FUNCTION "FRK_PersistCommitAnchor" : Void
{ S7_Optimized_Access := 'TRUE' }
VERSION : 0.1
VAR_INPUT
    Slot : Int;
END_VAR
BEGIN
    IF #Slot < 1 OR #Slot > 18 THEN RETURN; END_IF;
    IF "FRK_PersistAnchors".SelectedB[#Slot] THEN "FRK_PersistAnchors".RowsA[#Slot] := "FRK_PersistRuntime".Anchor[#Slot];
    ELSE "FRK_PersistAnchors".RowsB[#Slot] := "FRK_PersistRuntime".Anchor[#Slot]; END_IF;
    "FRK_PersistAnchors".SelectedB[#Slot] := NOT "FRK_PersistAnchors".SelectedB[#Slot];
    "FRK_PersistAnchors".Commissioned[#Slot] := TRUE;
END_FUNCTION
// Binding-owned byte medium. Consumers own content validation and authority.
FUNCTION "FRK_PersistNumber" : DWord
{ S7_Optimized_Access := 'TRUE' }
VERSION : 0.1
VAR_INPUT
    Offset : Int;
END_VAR
VAR_IN_OUT
    Bytes : Array[*] of Byte;
END_VAR
VAR_TEMP
    Index : Int;
END_VAR
BEGIN
    #FRK_PersistNumber := DWORD#0;
    IF #Offset < 0 OR #Offset > UPPER_BOUND(ARR := #Bytes, DIM := 1) - 3 THEN RETURN; END_IF;
    FOR #Index := 0 TO 3 DO
        #FRK_PersistNumber := #FRK_PersistNumber OR SHL(IN := BYTE_TO_DWORD(#Bytes[#Offset + #Index]), N := INT_TO_UINT(#Index * 8));
    END_FOR;
END_FUNCTION

FUNCTION "FRK_PersistPutNumber" : Void
{ S7_Optimized_Access := 'TRUE' }
VERSION : 0.1
VAR_INPUT
    Offset : Int;
    Value : DWord;
END_VAR
VAR_IN_OUT
    Bytes : Array[*] of Byte;
END_VAR
VAR_TEMP
    Index : Int;
END_VAR
BEGIN
    IF #Offset < 0 OR #Offset > UPPER_BOUND(ARR := #Bytes, DIM := 1) - 3 THEN RETURN; END_IF;
    FOR #Index := 0 TO 3 DO #Bytes[#Offset + #Index] := DWORD_TO_BYTE(SHR(IN := #Value, N := INT_TO_UINT(#Index * 8))); END_FOR;
END_FUNCTION

FUNCTION "FRK_PersistKeyCrc" : DWord
{ S7_Optimized_Access := 'TRUE' }
VERSION : 0.1
VAR_INPUT
    Key : String;
END_VAR
VAR_TEMP
    Index : Int;
    Work : DWord;
END_VAR
BEGIN
    #Work := "FRK_CrcNumber"(Previous := DWORD#16#FFFFFFFF, Value := INT_TO_UDINT(LEN(#Key)));
    FOR #Index := 1 TO LEN(#Key) DO #Work := "FRK_CrcByte"(Previous := #Work, Value := CHAR_TO_BYTE(#Key[#Index])); END_FOR;
    #FRK_PersistKeyCrc := NOT #Work;
END_FUNCTION

FUNCTION "FRK_PersistAnchorCrc" : DWord
{ S7_Optimized_Access := 'TRUE' }
VERSION : 0.1
VAR_IN_OUT
    Image : "FRK_PersistAnchor";
END_VAR
VAR_TEMP
    Work : DWord;
END_VAR
BEGIN
    #Work := "FRK_CrcNumber"(Previous := DWORD#16#FFFFFFFF, Value := UINT_TO_UDINT(#Image.SchemaVersion));
    #Work := "FRK_CrcNumber"(Previous := #Work, Value := DWORD_TO_UDINT(#Image.KeyCrc));
    #Work := "FRK_CrcNumber"(Previous := #Work, Value := #Image.Generation);
    #Work := "FRK_CrcNumber"(Previous := #Work, Value := DWORD_TO_UDINT(#Image.DocumentCrc));
    #FRK_PersistAnchorCrc := NOT #Work;
END_FUNCTION

FUNCTION "FRK_PersistAnchorValid" : Bool
{ S7_Optimized_Access := 'TRUE' }
VERSION : 0.1
VAR_INPUT
    Slot : Int;
END_VAR
BEGIN
    #FRK_PersistAnchorValid := FALSE;
    IF #Slot < 1 OR #Slot > 18 THEN RETURN; END_IF;
    #FRK_PersistAnchorValid := "FRK_PersistAnchors".Commissioned[#Slot]
        AND "FRK_PersistRuntime".Anchor[#Slot].SchemaVersion = 1
        AND "FRK_PersistRuntime".Anchor[#Slot].KeyCrc = "FRK_PersistRuntime".KeyCrc[#Slot]
        AND "FRK_PersistRuntime".Anchor[#Slot].Checksum = "FRK_PersistAnchorCrc"(Image := "FRK_PersistRuntime".Anchor[#Slot]);
END_FUNCTION

FUNCTION "FRK_PersistRepair" : Void
{ S7_Optimized_Access := 'TRUE' }
VERSION : 0.1
VAR_INPUT
    Slot : Int;
END_VAR
BEGIN
    // Trusted consumer seam; never a remote command or authorization authority.
    IF #Slot < 1 OR #Slot > 18 THEN RETURN; END_IF;
    IF NOT "FRK_PersistAnchorValid"(Slot := #Slot) THEN
        "FRK_PersistRuntime".Anchor[#Slot].SchemaVersion := 1;
        "FRK_PersistRuntime".Anchor[#Slot].KeyCrc := "FRK_PersistRuntime".KeyCrc[#Slot];
        "FRK_PersistRuntime".Anchor[#Slot].Generation := 0;
        "FRK_PersistRuntime".Anchor[#Slot].DocumentCrc := DWORD#0;
        "FRK_PersistRuntime".Anchor[#Slot].Checksum := "FRK_PersistAnchorCrc"(Image := "FRK_PersistRuntime".Anchor[#Slot]);
        "FRK_PersistAnchors".Commissioned[#Slot] := TRUE;
    END_IF;
    "FRK_PersistCommitAnchor"(Slot := #Slot);
END_FUNCTION

FUNCTION "FRK_PersistStart" : UDInt
{ S7_Optimized_Access := 'TRUE' }
VERSION : 0.1
VAR_INPUT
    Slot : Int;
    WriteDocument : Bool;
    Length : DInt;
END_VAR
VAR_TEMP
    Index : Int;
END_VAR
BEGIN
    #FRK_PersistStart := 0;
    IF #Slot < 1 OR #Slot > 18 THEN RETURN; END_IF;
    IF #Length < 0 OR #Length > "FRK_PersistRuntime".Capacity[#Slot] OR "FRK_PersistRuntime".Leased[#Slot] THEN RETURN; END_IF;
    IF "FRK_PersistRuntime".LastTicket = UDINT#4294967295 THEN RETURN; END_IF;
    FOR #Index := 1 TO 4 DO
        IF "FRK_PersistRuntime".Queue[#Index].State = 0 THEN
            "FRK_PersistRuntime".LastTicket := "FRK_PersistRuntime".LastTicket + 1;
            "FRK_PersistRuntime".Queue[#Index].Ticket := "FRK_PersistRuntime".LastTicket;
            "FRK_PersistRuntime".Queue[#Index].Slot := #Slot;
            "FRK_PersistRuntime".Queue[#Index].WriteDocument := #WriteDocument;
            "FRK_PersistRuntime".Queue[#Index].Length := #Length;
            "FRK_PersistRuntime".Queue[#Index].State := 1;
            "FRK_PersistRuntime".Leased[#Slot] := TRUE;
            #FRK_PersistStart := "FRK_PersistRuntime".LastTicket;
            RETURN;
        END_IF;
    END_FOR;
END_FUNCTION

FUNCTION "FRK_PersistFinish" : Void
{ S7_Optimized_Access := 'TRUE' }
VERSION : 0.1
BEGIN
    IF "FRK_PersistRuntime".Active < 1 OR "FRK_PersistRuntime".Active > 4 THEN RETURN; END_IF;
    "FRK_PersistRuntime".Queue["FRK_PersistRuntime".Active].Result := "FRK_PersistRuntime".Result;
    "FRK_PersistRuntime".Queue["FRK_PersistRuntime".Active].State := 3;
    "FRK_PersistRuntime".Active := 0;
    "FRK_PersistRuntime".Stage := 0;
END_FUNCTION

FUNCTION "FRK_PersistValidate" : Bool
{ S7_Optimized_Access := 'TRUE' }
VERSION : 0.1
VAR_INPUT
    ExpectedKey : DWord;
END_VAR
VAR_IN_OUT
    Bytes : Array[*] of Byte;
    Check : "FRK_PersistCheck";
END_VAR
VAR_TEMP
    Budget : Int;
    Offset : Int;
    Upper : Int;
END_VAR
BEGIN
    #FRK_PersistValidate := FALSE;
    #Upper := DINT_TO_INT(UPPER_BOUND(ARR := #Bytes, DIM := 1));
    IF #Check.Cursor = -1 THEN
        #Check.Valid := FALSE; #Check.Empty := TRUE; #Check.Generation := 0; #Check.Length := 0;
        #Check.Cursor := 0; #Check.Crc := DWORD#16#FFFFFFFF;
        #Check.ZeroMode := "FRK_PersistNumber"(Offset := 0, Bytes := #Bytes) = DWORD#0;
        IF NOT #Check.ZeroMode THEN
            #Check.Empty := FALSE;
            IF "FRK_PersistNumber"(Offset := 0, Bytes := #Bytes) <> DWORD#826559046
                OR "FRK_PersistNumber"(Offset := 4, Bytes := #Bytes) <> DWORD#1
                OR "FRK_PersistNumber"(Offset := 16, Bytes := #Bytes) <> #ExpectedKey THEN #FRK_PersistValidate := TRUE; RETURN; END_IF;
            #Check.Generation := DWORD_TO_UDINT("FRK_PersistNumber"(Offset := 8, Bytes := #Bytes));
            #Check.Length := DWORD_TO_UDINT("FRK_PersistNumber"(Offset := 12, Bytes := #Bytes));
            IF #Check.Generation = 0 OR #Check.Length > INT_TO_UDINT(#Upper + 1 - 24) THEN #FRK_PersistValidate := TRUE; RETURN; END_IF;
        END_IF;
    END_IF;
    #Budget := 0;
    IF #Check.ZeroMode THEN
        WHILE #Check.Cursor <= #Upper AND #Budget < 512 DO
            IF #Bytes[#Check.Cursor] <> BYTE#0 THEN #Check.Empty := FALSE; #FRK_PersistValidate := TRUE; RETURN; END_IF;
            #Check.Cursor := #Check.Cursor + 1; #Budget := #Budget + 1;
        END_WHILE;
        #FRK_PersistValidate := #Check.Cursor > #Upper;
    ELSE
        WHILE #Check.Cursor < 20 + UDINT_TO_DINT(#Check.Length) AND #Budget < 512 DO
            IF #Check.Cursor < 20 THEN #Offset := DINT_TO_INT(#Check.Cursor); ELSE #Offset := DINT_TO_INT(#Check.Cursor + 24 - 20); END_IF;
            #Check.Crc := "FRK_CrcByte"(Previous := #Check.Crc, Value := #Bytes[#Offset]);
            #Check.Cursor := #Check.Cursor + 1; #Budget := #Budget + 1;
        END_WHILE;
        IF #Check.Cursor >= 20 + UDINT_TO_DINT(#Check.Length) THEN
            #Check.Crc := NOT #Check.Crc;
            #Check.Valid := #Check.Crc = "FRK_PersistNumber"(Offset := 20, Bytes := #Bytes);
            #FRK_PersistValidate := TRUE;
        END_IF;
    END_IF;
END_FUNCTION

FUNCTION "FRK_PersistInspect" : Void
{ S7_Optimized_Access := 'TRUE' }
VERSION : 0.1
VAR_IN_OUT
    BytesA : Array[*] of Byte;
    BytesB : Array[*] of Byte;
    Payload : Array[*] of Byte;
END_VAR
VAR_TEMP
    Index : Int;
    Slot : Int;
    Chosen : Int;
    Generation : UDInt;
    Length : UDInt;
    DocumentCrc : DWord;
    Lost : Bool;
END_VAR
BEGIN
    #Slot := "FRK_PersistRuntime".Slot;
    #Chosen := 0; #Generation := 0; #Length := 0; #DocumentCrc := DWORD#0;
    IF "FRK_PersistRuntime".CheckA.Valid THEN
        #Chosen := 1; #Generation := "FRK_PersistRuntime".CheckA.Generation;
        #Length := "FRK_PersistRuntime".CheckA.Length; #DocumentCrc := "FRK_PersistRuntime".CheckA.Crc;
    END_IF;
    IF "FRK_PersistRuntime".CheckB.Valid AND (#Chosen = 0 OR "FRK_PersistRuntime".CheckB.Generation > #Generation) THEN
        #Chosen := 2; #Generation := "FRK_PersistRuntime".CheckB.Generation;
        #Length := "FRK_PersistRuntime".CheckB.Length; #DocumentCrc := "FRK_PersistRuntime".CheckB.Crc;
    END_IF;
    #Lost := #Generation < "FRK_PersistRuntime".Anchor[#Slot].Generation;
    IF "FRK_PersistRuntime".CheckA.Valid AND "FRK_PersistRuntime".CheckB.Valid
        AND "FRK_PersistRuntime".CheckA.Generation = "FRK_PersistRuntime".CheckB.Generation
        AND "FRK_PersistRuntime".CheckA.Crc <> "FRK_PersistRuntime".CheckB.Crc THEN #Chosen := 0; #Lost := TRUE; END_IF;
    IF #Chosen = 0 AND (NOT "FRK_PersistRuntime".CheckA.Empty OR NOT "FRK_PersistRuntime".CheckB.Empty) THEN #Lost := TRUE; END_IF;
    IF #Generation = "FRK_PersistRuntime".Anchor[#Slot].Generation AND #Generation > 0
        AND #DocumentCrc <> "FRK_PersistRuntime".Anchor[#Slot].DocumentCrc THEN #Chosen := 0; #Lost := TRUE; END_IF;
    IF NOT "FRK_PersistAnchorValid"(Slot := #Slot) THEN
        "FRK_PersistRuntime".Result.Lost := TRUE;
        IF "FRK_PersistRuntime".Queue["FRK_PersistRuntime".Active].WriteDocument THEN
            "FRK_PersistRuntime".Result.ErrorId := 2;
        ELSE "FRK_PersistRuntime".Result.Ok := TRUE; END_IF;
        "FRK_PersistFinish"(); RETURN;
    END_IF;
    IF NOT "FRK_PersistRuntime".Queue["FRK_PersistRuntime".Active].WriteDocument THEN
        "FRK_PersistRuntime".Result.Ok := TRUE;
        "FRK_PersistRuntime".Result.Lost := #Lost;
        "FRK_PersistRuntime".Result.Found := #Chosen <> 0 AND #Length > 0;
        "FRK_PersistRuntime".Result.Length := #Length;
        IF #Chosen = 0 THEN "FRK_PersistRuntime".Result.Length := 0; END_IF;
        IF #Chosen <> 0 THEN
            FOR #Index := 0 TO UDINT_TO_DINT(#Length) - 1 DO
                IF #Chosen = 1 THEN #Payload[24 + #Index] := #BytesA[24 + #Index];
                ELSE #Payload[24 + #Index] := #BytesB[24 + #Index]; END_IF;
            END_FOR;
        END_IF;
        "FRK_PersistFinish"(); RETURN;
    END_IF;
    #Generation := MAX(IN1 := #Generation, IN2 := "FRK_PersistRuntime".Anchor[#Slot].Generation);
    IF #Generation = UDINT#4294967295 THEN
        "FRK_PersistRuntime".Result.ErrorId := 3;
        "FRK_PersistFinish"(); RETURN;
    END_IF;
    "FRK_PersistRuntime".Generation := #Generation + 1;
    "FRK_PersistRuntime".Chosen := 2;
    IF #Chosen = 2 THEN "FRK_PersistRuntime".Chosen := 1; END_IF;
    "FRK_PersistPutNumber"(Bytes := #Payload, Offset := 0, Value := DWORD#826559046);
    "FRK_PersistPutNumber"(Bytes := #Payload, Offset := 4, Value := DWORD#1);
    "FRK_PersistPutNumber"(Bytes := #Payload, Offset := 8, Value := UDINT_TO_DWORD("FRK_PersistRuntime".Generation));
    "FRK_PersistPutNumber"(Bytes := #Payload, Offset := 12, Value := DINT_TO_DWORD("FRK_PersistRuntime".Queue["FRK_PersistRuntime".Active].Length));
    "FRK_PersistPutNumber"(Bytes := #Payload, Offset := 16, Value := "FRK_PersistRuntime".KeyCrc[#Slot]);
    "FRK_PersistRuntime".CheckWrite.Cursor := -1;
    "FRK_PersistRuntime".Stage := 6;
END_FUNCTION
FUNCTION "FRK_PersistIo" : Void
{ S7_Optimized_Access := 'TRUE' }
VERSION : 0.1
VAR_INPUT
    Operation : Int;
END_VAR
BEGIN
    CASE "FRK_PersistRuntime".Slot OF
        1:
            CASE #Operation OF
                1: "FRK_PersistRuntime".NativeResult := READ_DBL(REQ := "FRK_PersistRuntime".NativeReq, SRCBLK := "FRK_Load_D001A".Bytes, BUSY => "FRK_PersistRuntime".NativeBusy, DSTBLK => "FRK_PersistBuffers".D001A);
                2: "FRK_PersistRuntime".NativeResult := READ_DBL(REQ := "FRK_PersistRuntime".NativeReq, SRCBLK := "FRK_Load_D001B".Bytes, BUSY => "FRK_PersistRuntime".NativeBusy, DSTBLK => "FRK_PersistBuffers".D001B);
                3: "FRK_PersistRuntime".NativeResult := WRIT_DBL(REQ := "FRK_PersistRuntime".NativeReq, SRCBLK := "FRK_PersistBuffers".D001Data, BUSY => "FRK_PersistRuntime".NativeBusy, DSTBLK => "FRK_Load_D001A".Bytes);
                4: "FRK_PersistRuntime".NativeResult := WRIT_DBL(REQ := "FRK_PersistRuntime".NativeReq, SRCBLK := "FRK_PersistBuffers".D001Data, BUSY => "FRK_PersistRuntime".NativeBusy, DSTBLK => "FRK_Load_D001B".Bytes);
                ELSE "FRK_PersistRuntime".NativeResult := -1; "FRK_PersistRuntime".NativeBusy := FALSE;
            END_CASE;
        2:
            CASE #Operation OF
                1: "FRK_PersistRuntime".NativeResult := READ_DBL(REQ := "FRK_PersistRuntime".NativeReq, SRCBLK := "FRK_Load_D002A".Bytes, BUSY => "FRK_PersistRuntime".NativeBusy, DSTBLK => "FRK_PersistBuffers".D002A);
                2: "FRK_PersistRuntime".NativeResult := READ_DBL(REQ := "FRK_PersistRuntime".NativeReq, SRCBLK := "FRK_Load_D002B".Bytes, BUSY => "FRK_PersistRuntime".NativeBusy, DSTBLK => "FRK_PersistBuffers".D002B);
                3: "FRK_PersistRuntime".NativeResult := WRIT_DBL(REQ := "FRK_PersistRuntime".NativeReq, SRCBLK := "FRK_PersistBuffers".D002Data, BUSY => "FRK_PersistRuntime".NativeBusy, DSTBLK => "FRK_Load_D002A".Bytes);
                4: "FRK_PersistRuntime".NativeResult := WRIT_DBL(REQ := "FRK_PersistRuntime".NativeReq, SRCBLK := "FRK_PersistBuffers".D002Data, BUSY => "FRK_PersistRuntime".NativeBusy, DSTBLK => "FRK_Load_D002B".Bytes);
                ELSE "FRK_PersistRuntime".NativeResult := -1; "FRK_PersistRuntime".NativeBusy := FALSE;
            END_CASE;
        3:
            CASE #Operation OF
                1: "FRK_PersistRuntime".NativeResult := READ_DBL(REQ := "FRK_PersistRuntime".NativeReq, SRCBLK := "FRK_Load_D003A".Bytes, BUSY => "FRK_PersistRuntime".NativeBusy, DSTBLK => "FRK_PersistBuffers".D003A);
                2: "FRK_PersistRuntime".NativeResult := READ_DBL(REQ := "FRK_PersistRuntime".NativeReq, SRCBLK := "FRK_Load_D003B".Bytes, BUSY => "FRK_PersistRuntime".NativeBusy, DSTBLK => "FRK_PersistBuffers".D003B);
                3: "FRK_PersistRuntime".NativeResult := WRIT_DBL(REQ := "FRK_PersistRuntime".NativeReq, SRCBLK := "FRK_PersistBuffers".D003Data, BUSY => "FRK_PersistRuntime".NativeBusy, DSTBLK => "FRK_Load_D003A".Bytes);
                4: "FRK_PersistRuntime".NativeResult := WRIT_DBL(REQ := "FRK_PersistRuntime".NativeReq, SRCBLK := "FRK_PersistBuffers".D003Data, BUSY => "FRK_PersistRuntime".NativeBusy, DSTBLK => "FRK_Load_D003B".Bytes);
                ELSE "FRK_PersistRuntime".NativeResult := -1; "FRK_PersistRuntime".NativeBusy := FALSE;
            END_CASE;
        4:
            CASE #Operation OF
                1: "FRK_PersistRuntime".NativeResult := READ_DBL(REQ := "FRK_PersistRuntime".NativeReq, SRCBLK := "FRK_Load_D004A".Bytes, BUSY => "FRK_PersistRuntime".NativeBusy, DSTBLK => "FRK_PersistBuffers".D004A);
                2: "FRK_PersistRuntime".NativeResult := READ_DBL(REQ := "FRK_PersistRuntime".NativeReq, SRCBLK := "FRK_Load_D004B".Bytes, BUSY => "FRK_PersistRuntime".NativeBusy, DSTBLK => "FRK_PersistBuffers".D004B);
                3: "FRK_PersistRuntime".NativeResult := WRIT_DBL(REQ := "FRK_PersistRuntime".NativeReq, SRCBLK := "FRK_PersistBuffers".D004Data, BUSY => "FRK_PersistRuntime".NativeBusy, DSTBLK => "FRK_Load_D004A".Bytes);
                4: "FRK_PersistRuntime".NativeResult := WRIT_DBL(REQ := "FRK_PersistRuntime".NativeReq, SRCBLK := "FRK_PersistBuffers".D004Data, BUSY => "FRK_PersistRuntime".NativeBusy, DSTBLK => "FRK_Load_D004B".Bytes);
                ELSE "FRK_PersistRuntime".NativeResult := -1; "FRK_PersistRuntime".NativeBusy := FALSE;
            END_CASE;
        5:
            CASE #Operation OF
                1: "FRK_PersistRuntime".NativeResult := READ_DBL(REQ := "FRK_PersistRuntime".NativeReq, SRCBLK := "FRK_Load_D005A".Bytes, BUSY => "FRK_PersistRuntime".NativeBusy, DSTBLK => "FRK_PersistBuffers".D005A);
                2: "FRK_PersistRuntime".NativeResult := READ_DBL(REQ := "FRK_PersistRuntime".NativeReq, SRCBLK := "FRK_Load_D005B".Bytes, BUSY => "FRK_PersistRuntime".NativeBusy, DSTBLK => "FRK_PersistBuffers".D005B);
                3: "FRK_PersistRuntime".NativeResult := WRIT_DBL(REQ := "FRK_PersistRuntime".NativeReq, SRCBLK := "FRK_PersistBuffers".D005Data, BUSY => "FRK_PersistRuntime".NativeBusy, DSTBLK => "FRK_Load_D005A".Bytes);
                4: "FRK_PersistRuntime".NativeResult := WRIT_DBL(REQ := "FRK_PersistRuntime".NativeReq, SRCBLK := "FRK_PersistBuffers".D005Data, BUSY => "FRK_PersistRuntime".NativeBusy, DSTBLK => "FRK_Load_D005B".Bytes);
                ELSE "FRK_PersistRuntime".NativeResult := -1; "FRK_PersistRuntime".NativeBusy := FALSE;
            END_CASE;
        6:
            CASE #Operation OF
                1: "FRK_PersistRuntime".NativeResult := READ_DBL(REQ := "FRK_PersistRuntime".NativeReq, SRCBLK := "FRK_Load_D006A".Bytes, BUSY => "FRK_PersistRuntime".NativeBusy, DSTBLK => "FRK_PersistBuffers".D006A);
                2: "FRK_PersistRuntime".NativeResult := READ_DBL(REQ := "FRK_PersistRuntime".NativeReq, SRCBLK := "FRK_Load_D006B".Bytes, BUSY => "FRK_PersistRuntime".NativeBusy, DSTBLK => "FRK_PersistBuffers".D006B);
                3: "FRK_PersistRuntime".NativeResult := WRIT_DBL(REQ := "FRK_PersistRuntime".NativeReq, SRCBLK := "FRK_PersistBuffers".D006Data, BUSY => "FRK_PersistRuntime".NativeBusy, DSTBLK => "FRK_Load_D006A".Bytes);
                4: "FRK_PersistRuntime".NativeResult := WRIT_DBL(REQ := "FRK_PersistRuntime".NativeReq, SRCBLK := "FRK_PersistBuffers".D006Data, BUSY => "FRK_PersistRuntime".NativeBusy, DSTBLK => "FRK_Load_D006B".Bytes);
                ELSE "FRK_PersistRuntime".NativeResult := -1; "FRK_PersistRuntime".NativeBusy := FALSE;
            END_CASE;
        7:
            CASE #Operation OF
                1: "FRK_PersistRuntime".NativeResult := READ_DBL(REQ := "FRK_PersistRuntime".NativeReq, SRCBLK := "FRK_Load_D007A".Bytes, BUSY => "FRK_PersistRuntime".NativeBusy, DSTBLK => "FRK_PersistBuffers".D007A);
                2: "FRK_PersistRuntime".NativeResult := READ_DBL(REQ := "FRK_PersistRuntime".NativeReq, SRCBLK := "FRK_Load_D007B".Bytes, BUSY => "FRK_PersistRuntime".NativeBusy, DSTBLK => "FRK_PersistBuffers".D007B);
                3: "FRK_PersistRuntime".NativeResult := WRIT_DBL(REQ := "FRK_PersistRuntime".NativeReq, SRCBLK := "FRK_PersistBuffers".D007Data, BUSY => "FRK_PersistRuntime".NativeBusy, DSTBLK => "FRK_Load_D007A".Bytes);
                4: "FRK_PersistRuntime".NativeResult := WRIT_DBL(REQ := "FRK_PersistRuntime".NativeReq, SRCBLK := "FRK_PersistBuffers".D007Data, BUSY => "FRK_PersistRuntime".NativeBusy, DSTBLK => "FRK_Load_D007B".Bytes);
                ELSE "FRK_PersistRuntime".NativeResult := -1; "FRK_PersistRuntime".NativeBusy := FALSE;
            END_CASE;
        8:
            CASE #Operation OF
                1: "FRK_PersistRuntime".NativeResult := READ_DBL(REQ := "FRK_PersistRuntime".NativeReq, SRCBLK := "FRK_Load_D008A".Bytes, BUSY => "FRK_PersistRuntime".NativeBusy, DSTBLK => "FRK_PersistBuffers".D008A);
                2: "FRK_PersistRuntime".NativeResult := READ_DBL(REQ := "FRK_PersistRuntime".NativeReq, SRCBLK := "FRK_Load_D008B".Bytes, BUSY => "FRK_PersistRuntime".NativeBusy, DSTBLK => "FRK_PersistBuffers".D008B);
                3: "FRK_PersistRuntime".NativeResult := WRIT_DBL(REQ := "FRK_PersistRuntime".NativeReq, SRCBLK := "FRK_PersistBuffers".D008Data, BUSY => "FRK_PersistRuntime".NativeBusy, DSTBLK => "FRK_Load_D008A".Bytes);
                4: "FRK_PersistRuntime".NativeResult := WRIT_DBL(REQ := "FRK_PersistRuntime".NativeReq, SRCBLK := "FRK_PersistBuffers".D008Data, BUSY => "FRK_PersistRuntime".NativeBusy, DSTBLK => "FRK_Load_D008B".Bytes);
                ELSE "FRK_PersistRuntime".NativeResult := -1; "FRK_PersistRuntime".NativeBusy := FALSE;
            END_CASE;
        9:
            CASE #Operation OF
                1: "FRK_PersistRuntime".NativeResult := READ_DBL(REQ := "FRK_PersistRuntime".NativeReq, SRCBLK := "FRK_Load_D009A".Bytes, BUSY => "FRK_PersistRuntime".NativeBusy, DSTBLK => "FRK_PersistBuffers".D009A);
                2: "FRK_PersistRuntime".NativeResult := READ_DBL(REQ := "FRK_PersistRuntime".NativeReq, SRCBLK := "FRK_Load_D009B".Bytes, BUSY => "FRK_PersistRuntime".NativeBusy, DSTBLK => "FRK_PersistBuffers".D009B);
                3: "FRK_PersistRuntime".NativeResult := WRIT_DBL(REQ := "FRK_PersistRuntime".NativeReq, SRCBLK := "FRK_PersistBuffers".D009Data, BUSY => "FRK_PersistRuntime".NativeBusy, DSTBLK => "FRK_Load_D009A".Bytes);
                4: "FRK_PersistRuntime".NativeResult := WRIT_DBL(REQ := "FRK_PersistRuntime".NativeReq, SRCBLK := "FRK_PersistBuffers".D009Data, BUSY => "FRK_PersistRuntime".NativeBusy, DSTBLK => "FRK_Load_D009B".Bytes);
                ELSE "FRK_PersistRuntime".NativeResult := -1; "FRK_PersistRuntime".NativeBusy := FALSE;
            END_CASE;
        10:
            CASE #Operation OF
                1: "FRK_PersistRuntime".NativeResult := READ_DBL(REQ := "FRK_PersistRuntime".NativeReq, SRCBLK := "FRK_Load_D010A".Bytes, BUSY => "FRK_PersistRuntime".NativeBusy, DSTBLK => "FRK_PersistBuffers".D010A);
                2: "FRK_PersistRuntime".NativeResult := READ_DBL(REQ := "FRK_PersistRuntime".NativeReq, SRCBLK := "FRK_Load_D010B".Bytes, BUSY => "FRK_PersistRuntime".NativeBusy, DSTBLK => "FRK_PersistBuffers".D010B);
                3: "FRK_PersistRuntime".NativeResult := WRIT_DBL(REQ := "FRK_PersistRuntime".NativeReq, SRCBLK := "FRK_PersistBuffers".D010Data, BUSY => "FRK_PersistRuntime".NativeBusy, DSTBLK => "FRK_Load_D010A".Bytes);
                4: "FRK_PersistRuntime".NativeResult := WRIT_DBL(REQ := "FRK_PersistRuntime".NativeReq, SRCBLK := "FRK_PersistBuffers".D010Data, BUSY => "FRK_PersistRuntime".NativeBusy, DSTBLK => "FRK_Load_D010B".Bytes);
                ELSE "FRK_PersistRuntime".NativeResult := -1; "FRK_PersistRuntime".NativeBusy := FALSE;
            END_CASE;
        11:
            CASE #Operation OF
                1: "FRK_PersistRuntime".NativeResult := READ_DBL(REQ := "FRK_PersistRuntime".NativeReq, SRCBLK := "FRK_Load_D011A".Bytes, BUSY => "FRK_PersistRuntime".NativeBusy, DSTBLK => "FRK_PersistBuffers".D011A);
                2: "FRK_PersistRuntime".NativeResult := READ_DBL(REQ := "FRK_PersistRuntime".NativeReq, SRCBLK := "FRK_Load_D011B".Bytes, BUSY => "FRK_PersistRuntime".NativeBusy, DSTBLK => "FRK_PersistBuffers".D011B);
                3: "FRK_PersistRuntime".NativeResult := WRIT_DBL(REQ := "FRK_PersistRuntime".NativeReq, SRCBLK := "FRK_PersistBuffers".D011Data, BUSY => "FRK_PersistRuntime".NativeBusy, DSTBLK => "FRK_Load_D011A".Bytes);
                4: "FRK_PersistRuntime".NativeResult := WRIT_DBL(REQ := "FRK_PersistRuntime".NativeReq, SRCBLK := "FRK_PersistBuffers".D011Data, BUSY => "FRK_PersistRuntime".NativeBusy, DSTBLK => "FRK_Load_D011B".Bytes);
                ELSE "FRK_PersistRuntime".NativeResult := -1; "FRK_PersistRuntime".NativeBusy := FALSE;
            END_CASE;
        12:
            CASE #Operation OF
                1: "FRK_PersistRuntime".NativeResult := READ_DBL(REQ := "FRK_PersistRuntime".NativeReq, SRCBLK := "FRK_Load_D012A".Bytes, BUSY => "FRK_PersistRuntime".NativeBusy, DSTBLK => "FRK_PersistBuffers".D012A);
                2: "FRK_PersistRuntime".NativeResult := READ_DBL(REQ := "FRK_PersistRuntime".NativeReq, SRCBLK := "FRK_Load_D012B".Bytes, BUSY => "FRK_PersistRuntime".NativeBusy, DSTBLK => "FRK_PersistBuffers".D012B);
                3: "FRK_PersistRuntime".NativeResult := WRIT_DBL(REQ := "FRK_PersistRuntime".NativeReq, SRCBLK := "FRK_PersistBuffers".D012Data, BUSY => "FRK_PersistRuntime".NativeBusy, DSTBLK => "FRK_Load_D012A".Bytes);
                4: "FRK_PersistRuntime".NativeResult := WRIT_DBL(REQ := "FRK_PersistRuntime".NativeReq, SRCBLK := "FRK_PersistBuffers".D012Data, BUSY => "FRK_PersistRuntime".NativeBusy, DSTBLK => "FRK_Load_D012B".Bytes);
                ELSE "FRK_PersistRuntime".NativeResult := -1; "FRK_PersistRuntime".NativeBusy := FALSE;
            END_CASE;
        13:
            CASE #Operation OF
                1: "FRK_PersistRuntime".NativeResult := READ_DBL(REQ := "FRK_PersistRuntime".NativeReq, SRCBLK := "FRK_Load_D013A".Bytes, BUSY => "FRK_PersistRuntime".NativeBusy, DSTBLK => "FRK_PersistBuffers".D013A);
                2: "FRK_PersistRuntime".NativeResult := READ_DBL(REQ := "FRK_PersistRuntime".NativeReq, SRCBLK := "FRK_Load_D013B".Bytes, BUSY => "FRK_PersistRuntime".NativeBusy, DSTBLK => "FRK_PersistBuffers".D013B);
                3: "FRK_PersistRuntime".NativeResult := WRIT_DBL(REQ := "FRK_PersistRuntime".NativeReq, SRCBLK := "FRK_PersistBuffers".D013Data, BUSY => "FRK_PersistRuntime".NativeBusy, DSTBLK => "FRK_Load_D013A".Bytes);
                4: "FRK_PersistRuntime".NativeResult := WRIT_DBL(REQ := "FRK_PersistRuntime".NativeReq, SRCBLK := "FRK_PersistBuffers".D013Data, BUSY => "FRK_PersistRuntime".NativeBusy, DSTBLK => "FRK_Load_D013B".Bytes);
                ELSE "FRK_PersistRuntime".NativeResult := -1; "FRK_PersistRuntime".NativeBusy := FALSE;
            END_CASE;
        14:
            CASE #Operation OF
                1: "FRK_PersistRuntime".NativeResult := READ_DBL(REQ := "FRK_PersistRuntime".NativeReq, SRCBLK := "FRK_Load_D014A".Bytes, BUSY => "FRK_PersistRuntime".NativeBusy, DSTBLK => "FRK_PersistBuffers".D014A);
                2: "FRK_PersistRuntime".NativeResult := READ_DBL(REQ := "FRK_PersistRuntime".NativeReq, SRCBLK := "FRK_Load_D014B".Bytes, BUSY => "FRK_PersistRuntime".NativeBusy, DSTBLK => "FRK_PersistBuffers".D014B);
                3: "FRK_PersistRuntime".NativeResult := WRIT_DBL(REQ := "FRK_PersistRuntime".NativeReq, SRCBLK := "FRK_PersistBuffers".D014Data, BUSY => "FRK_PersistRuntime".NativeBusy, DSTBLK => "FRK_Load_D014A".Bytes);
                4: "FRK_PersistRuntime".NativeResult := WRIT_DBL(REQ := "FRK_PersistRuntime".NativeReq, SRCBLK := "FRK_PersistBuffers".D014Data, BUSY => "FRK_PersistRuntime".NativeBusy, DSTBLK => "FRK_Load_D014B".Bytes);
                ELSE "FRK_PersistRuntime".NativeResult := -1; "FRK_PersistRuntime".NativeBusy := FALSE;
            END_CASE;
        15:
            CASE #Operation OF
                1: "FRK_PersistRuntime".NativeResult := READ_DBL(REQ := "FRK_PersistRuntime".NativeReq, SRCBLK := "FRK_Load_D015A".Bytes, BUSY => "FRK_PersistRuntime".NativeBusy, DSTBLK => "FRK_PersistBuffers".D015A);
                2: "FRK_PersistRuntime".NativeResult := READ_DBL(REQ := "FRK_PersistRuntime".NativeReq, SRCBLK := "FRK_Load_D015B".Bytes, BUSY => "FRK_PersistRuntime".NativeBusy, DSTBLK => "FRK_PersistBuffers".D015B);
                3: "FRK_PersistRuntime".NativeResult := WRIT_DBL(REQ := "FRK_PersistRuntime".NativeReq, SRCBLK := "FRK_PersistBuffers".D015Data, BUSY => "FRK_PersistRuntime".NativeBusy, DSTBLK => "FRK_Load_D015A".Bytes);
                4: "FRK_PersistRuntime".NativeResult := WRIT_DBL(REQ := "FRK_PersistRuntime".NativeReq, SRCBLK := "FRK_PersistBuffers".D015Data, BUSY => "FRK_PersistRuntime".NativeBusy, DSTBLK => "FRK_Load_D015B".Bytes);
                ELSE "FRK_PersistRuntime".NativeResult := -1; "FRK_PersistRuntime".NativeBusy := FALSE;
            END_CASE;
        16:
            CASE #Operation OF
                1: "FRK_PersistRuntime".NativeResult := READ_DBL(REQ := "FRK_PersistRuntime".NativeReq, SRCBLK := "FRK_Load_D016A".Bytes, BUSY => "FRK_PersistRuntime".NativeBusy, DSTBLK => "FRK_PersistBuffers".D016A);
                2: "FRK_PersistRuntime".NativeResult := READ_DBL(REQ := "FRK_PersistRuntime".NativeReq, SRCBLK := "FRK_Load_D016B".Bytes, BUSY => "FRK_PersistRuntime".NativeBusy, DSTBLK => "FRK_PersistBuffers".D016B);
                3: "FRK_PersistRuntime".NativeResult := WRIT_DBL(REQ := "FRK_PersistRuntime".NativeReq, SRCBLK := "FRK_PersistBuffers".D016Data, BUSY => "FRK_PersistRuntime".NativeBusy, DSTBLK => "FRK_Load_D016A".Bytes);
                4: "FRK_PersistRuntime".NativeResult := WRIT_DBL(REQ := "FRK_PersistRuntime".NativeReq, SRCBLK := "FRK_PersistBuffers".D016Data, BUSY => "FRK_PersistRuntime".NativeBusy, DSTBLK => "FRK_Load_D016B".Bytes);
                ELSE "FRK_PersistRuntime".NativeResult := -1; "FRK_PersistRuntime".NativeBusy := FALSE;
            END_CASE;
        17:
            CASE #Operation OF
                1: "FRK_PersistRuntime".NativeResult := READ_DBL(REQ := "FRK_PersistRuntime".NativeReq, SRCBLK := "FRK_Load_D017A".Bytes, BUSY => "FRK_PersistRuntime".NativeBusy, DSTBLK => "FRK_PersistBuffers".D017A);
                2: "FRK_PersistRuntime".NativeResult := READ_DBL(REQ := "FRK_PersistRuntime".NativeReq, SRCBLK := "FRK_Load_D017B".Bytes, BUSY => "FRK_PersistRuntime".NativeBusy, DSTBLK => "FRK_PersistBuffers".D017B);
                3: "FRK_PersistRuntime".NativeResult := WRIT_DBL(REQ := "FRK_PersistRuntime".NativeReq, SRCBLK := "FRK_PersistBuffers".D017Data, BUSY => "FRK_PersistRuntime".NativeBusy, DSTBLK => "FRK_Load_D017A".Bytes);
                4: "FRK_PersistRuntime".NativeResult := WRIT_DBL(REQ := "FRK_PersistRuntime".NativeReq, SRCBLK := "FRK_PersistBuffers".D017Data, BUSY => "FRK_PersistRuntime".NativeBusy, DSTBLK => "FRK_Load_D017B".Bytes);
                ELSE "FRK_PersistRuntime".NativeResult := -1; "FRK_PersistRuntime".NativeBusy := FALSE;
            END_CASE;
        18:
            CASE #Operation OF
                1: "FRK_PersistRuntime".NativeResult := READ_DBL(REQ := "FRK_PersistRuntime".NativeReq, SRCBLK := "FRK_Load_D018A".Bytes, BUSY => "FRK_PersistRuntime".NativeBusy, DSTBLK => "FRK_PersistBuffers".D018A);
                2: "FRK_PersistRuntime".NativeResult := READ_DBL(REQ := "FRK_PersistRuntime".NativeReq, SRCBLK := "FRK_Load_D018B".Bytes, BUSY => "FRK_PersistRuntime".NativeBusy, DSTBLK => "FRK_PersistBuffers".D018B);
                3: "FRK_PersistRuntime".NativeResult := WRIT_DBL(REQ := "FRK_PersistRuntime".NativeReq, SRCBLK := "FRK_PersistBuffers".D018Data, BUSY => "FRK_PersistRuntime".NativeBusy, DSTBLK => "FRK_Load_D018A".Bytes);
                4: "FRK_PersistRuntime".NativeResult := WRIT_DBL(REQ := "FRK_PersistRuntime".NativeReq, SRCBLK := "FRK_PersistBuffers".D018Data, BUSY => "FRK_PersistRuntime".NativeBusy, DSTBLK => "FRK_Load_D018B".Bytes);
                ELSE "FRK_PersistRuntime".NativeResult := -1; "FRK_PersistRuntime".NativeBusy := FALSE;
            END_CASE;
        ELSE "FRK_PersistRuntime".NativeResult := -1; "FRK_PersistRuntime".NativeBusy := FALSE;
    END_CASE;
END_FUNCTION
FUNCTION "FRK_PersistCheckA" : Bool
{ S7_Optimized_Access := 'TRUE' }
VERSION : 0.1
VAR_TEMP
    Done : Bool;
END_VAR
BEGIN
    #Done := FALSE;
    #FRK_PersistCheckA := FALSE;
    CASE "FRK_PersistRuntime".Slot OF
        1: #Done := "FRK_PersistValidate"(ExpectedKey := "FRK_PersistRuntime".KeyCrc[1], Bytes := "FRK_PersistBuffers".D001A, Check := "FRK_PersistRuntime".CheckA);
        2: #Done := "FRK_PersistValidate"(ExpectedKey := "FRK_PersistRuntime".KeyCrc[2], Bytes := "FRK_PersistBuffers".D002A, Check := "FRK_PersistRuntime".CheckA);
        3: #Done := "FRK_PersistValidate"(ExpectedKey := "FRK_PersistRuntime".KeyCrc[3], Bytes := "FRK_PersistBuffers".D003A, Check := "FRK_PersistRuntime".CheckA);
        4: #Done := "FRK_PersistValidate"(ExpectedKey := "FRK_PersistRuntime".KeyCrc[4], Bytes := "FRK_PersistBuffers".D004A, Check := "FRK_PersistRuntime".CheckA);
        5: #Done := "FRK_PersistValidate"(ExpectedKey := "FRK_PersistRuntime".KeyCrc[5], Bytes := "FRK_PersistBuffers".D005A, Check := "FRK_PersistRuntime".CheckA);
        6: #Done := "FRK_PersistValidate"(ExpectedKey := "FRK_PersistRuntime".KeyCrc[6], Bytes := "FRK_PersistBuffers".D006A, Check := "FRK_PersistRuntime".CheckA);
        7: #Done := "FRK_PersistValidate"(ExpectedKey := "FRK_PersistRuntime".KeyCrc[7], Bytes := "FRK_PersistBuffers".D007A, Check := "FRK_PersistRuntime".CheckA);
        8: #Done := "FRK_PersistValidate"(ExpectedKey := "FRK_PersistRuntime".KeyCrc[8], Bytes := "FRK_PersistBuffers".D008A, Check := "FRK_PersistRuntime".CheckA);
        9: #Done := "FRK_PersistValidate"(ExpectedKey := "FRK_PersistRuntime".KeyCrc[9], Bytes := "FRK_PersistBuffers".D009A, Check := "FRK_PersistRuntime".CheckA);
        10: #Done := "FRK_PersistValidate"(ExpectedKey := "FRK_PersistRuntime".KeyCrc[10], Bytes := "FRK_PersistBuffers".D010A, Check := "FRK_PersistRuntime".CheckA);
        11: #Done := "FRK_PersistValidate"(ExpectedKey := "FRK_PersistRuntime".KeyCrc[11], Bytes := "FRK_PersistBuffers".D011A, Check := "FRK_PersistRuntime".CheckA);
        12: #Done := "FRK_PersistValidate"(ExpectedKey := "FRK_PersistRuntime".KeyCrc[12], Bytes := "FRK_PersistBuffers".D012A, Check := "FRK_PersistRuntime".CheckA);
        13: #Done := "FRK_PersistValidate"(ExpectedKey := "FRK_PersistRuntime".KeyCrc[13], Bytes := "FRK_PersistBuffers".D013A, Check := "FRK_PersistRuntime".CheckA);
        14: #Done := "FRK_PersistValidate"(ExpectedKey := "FRK_PersistRuntime".KeyCrc[14], Bytes := "FRK_PersistBuffers".D014A, Check := "FRK_PersistRuntime".CheckA);
        15: #Done := "FRK_PersistValidate"(ExpectedKey := "FRK_PersistRuntime".KeyCrc[15], Bytes := "FRK_PersistBuffers".D015A, Check := "FRK_PersistRuntime".CheckA);
        16: #Done := "FRK_PersistValidate"(ExpectedKey := "FRK_PersistRuntime".KeyCrc[16], Bytes := "FRK_PersistBuffers".D016A, Check := "FRK_PersistRuntime".CheckA);
        17: #Done := "FRK_PersistValidate"(ExpectedKey := "FRK_PersistRuntime".KeyCrc[17], Bytes := "FRK_PersistBuffers".D017A, Check := "FRK_PersistRuntime".CheckA);
        18: #Done := "FRK_PersistValidate"(ExpectedKey := "FRK_PersistRuntime".KeyCrc[18], Bytes := "FRK_PersistBuffers".D018A, Check := "FRK_PersistRuntime".CheckA);
        ELSE RETURN;
    END_CASE;
    #FRK_PersistCheckA := #Done;
END_FUNCTION
FUNCTION "FRK_PersistCheckB" : Bool
{ S7_Optimized_Access := 'TRUE' }
VERSION : 0.1
VAR_TEMP
    Done : Bool;
END_VAR
BEGIN
    #Done := FALSE;
    #FRK_PersistCheckB := FALSE;
    CASE "FRK_PersistRuntime".Slot OF
        1: #Done := "FRK_PersistValidate"(ExpectedKey := "FRK_PersistRuntime".KeyCrc[1], Bytes := "FRK_PersistBuffers".D001B, Check := "FRK_PersistRuntime".CheckB);
        2: #Done := "FRK_PersistValidate"(ExpectedKey := "FRK_PersistRuntime".KeyCrc[2], Bytes := "FRK_PersistBuffers".D002B, Check := "FRK_PersistRuntime".CheckB);
        3: #Done := "FRK_PersistValidate"(ExpectedKey := "FRK_PersistRuntime".KeyCrc[3], Bytes := "FRK_PersistBuffers".D003B, Check := "FRK_PersistRuntime".CheckB);
        4: #Done := "FRK_PersistValidate"(ExpectedKey := "FRK_PersistRuntime".KeyCrc[4], Bytes := "FRK_PersistBuffers".D004B, Check := "FRK_PersistRuntime".CheckB);
        5: #Done := "FRK_PersistValidate"(ExpectedKey := "FRK_PersistRuntime".KeyCrc[5], Bytes := "FRK_PersistBuffers".D005B, Check := "FRK_PersistRuntime".CheckB);
        6: #Done := "FRK_PersistValidate"(ExpectedKey := "FRK_PersistRuntime".KeyCrc[6], Bytes := "FRK_PersistBuffers".D006B, Check := "FRK_PersistRuntime".CheckB);
        7: #Done := "FRK_PersistValidate"(ExpectedKey := "FRK_PersistRuntime".KeyCrc[7], Bytes := "FRK_PersistBuffers".D007B, Check := "FRK_PersistRuntime".CheckB);
        8: #Done := "FRK_PersistValidate"(ExpectedKey := "FRK_PersistRuntime".KeyCrc[8], Bytes := "FRK_PersistBuffers".D008B, Check := "FRK_PersistRuntime".CheckB);
        9: #Done := "FRK_PersistValidate"(ExpectedKey := "FRK_PersistRuntime".KeyCrc[9], Bytes := "FRK_PersistBuffers".D009B, Check := "FRK_PersistRuntime".CheckB);
        10: #Done := "FRK_PersistValidate"(ExpectedKey := "FRK_PersistRuntime".KeyCrc[10], Bytes := "FRK_PersistBuffers".D010B, Check := "FRK_PersistRuntime".CheckB);
        11: #Done := "FRK_PersistValidate"(ExpectedKey := "FRK_PersistRuntime".KeyCrc[11], Bytes := "FRK_PersistBuffers".D011B, Check := "FRK_PersistRuntime".CheckB);
        12: #Done := "FRK_PersistValidate"(ExpectedKey := "FRK_PersistRuntime".KeyCrc[12], Bytes := "FRK_PersistBuffers".D012B, Check := "FRK_PersistRuntime".CheckB);
        13: #Done := "FRK_PersistValidate"(ExpectedKey := "FRK_PersistRuntime".KeyCrc[13], Bytes := "FRK_PersistBuffers".D013B, Check := "FRK_PersistRuntime".CheckB);
        14: #Done := "FRK_PersistValidate"(ExpectedKey := "FRK_PersistRuntime".KeyCrc[14], Bytes := "FRK_PersistBuffers".D014B, Check := "FRK_PersistRuntime".CheckB);
        15: #Done := "FRK_PersistValidate"(ExpectedKey := "FRK_PersistRuntime".KeyCrc[15], Bytes := "FRK_PersistBuffers".D015B, Check := "FRK_PersistRuntime".CheckB);
        16: #Done := "FRK_PersistValidate"(ExpectedKey := "FRK_PersistRuntime".KeyCrc[16], Bytes := "FRK_PersistBuffers".D016B, Check := "FRK_PersistRuntime".CheckB);
        17: #Done := "FRK_PersistValidate"(ExpectedKey := "FRK_PersistRuntime".KeyCrc[17], Bytes := "FRK_PersistBuffers".D017B, Check := "FRK_PersistRuntime".CheckB);
        18: #Done := "FRK_PersistValidate"(ExpectedKey := "FRK_PersistRuntime".KeyCrc[18], Bytes := "FRK_PersistBuffers".D018B, Check := "FRK_PersistRuntime".CheckB);
        ELSE RETURN;
    END_CASE;
    #FRK_PersistCheckB := #Done;
END_FUNCTION
FUNCTION "FRK_PersistCheckWrite" : Bool
{ S7_Optimized_Access := 'TRUE' }
VERSION : 0.1
VAR_TEMP
    Done : Bool;
END_VAR
BEGIN
    #Done := FALSE;
    #FRK_PersistCheckWrite := FALSE;
    CASE "FRK_PersistRuntime".Slot OF
        1: #Done := "FRK_PersistValidate"(ExpectedKey := "FRK_PersistRuntime".KeyCrc[1], Bytes := "FRK_PersistBuffers".D001Data, Check := "FRK_PersistRuntime".CheckWrite);
        2: #Done := "FRK_PersistValidate"(ExpectedKey := "FRK_PersistRuntime".KeyCrc[2], Bytes := "FRK_PersistBuffers".D002Data, Check := "FRK_PersistRuntime".CheckWrite);
        3: #Done := "FRK_PersistValidate"(ExpectedKey := "FRK_PersistRuntime".KeyCrc[3], Bytes := "FRK_PersistBuffers".D003Data, Check := "FRK_PersistRuntime".CheckWrite);
        4: #Done := "FRK_PersistValidate"(ExpectedKey := "FRK_PersistRuntime".KeyCrc[4], Bytes := "FRK_PersistBuffers".D004Data, Check := "FRK_PersistRuntime".CheckWrite);
        5: #Done := "FRK_PersistValidate"(ExpectedKey := "FRK_PersistRuntime".KeyCrc[5], Bytes := "FRK_PersistBuffers".D005Data, Check := "FRK_PersistRuntime".CheckWrite);
        6: #Done := "FRK_PersistValidate"(ExpectedKey := "FRK_PersistRuntime".KeyCrc[6], Bytes := "FRK_PersistBuffers".D006Data, Check := "FRK_PersistRuntime".CheckWrite);
        7: #Done := "FRK_PersistValidate"(ExpectedKey := "FRK_PersistRuntime".KeyCrc[7], Bytes := "FRK_PersistBuffers".D007Data, Check := "FRK_PersistRuntime".CheckWrite);
        8: #Done := "FRK_PersistValidate"(ExpectedKey := "FRK_PersistRuntime".KeyCrc[8], Bytes := "FRK_PersistBuffers".D008Data, Check := "FRK_PersistRuntime".CheckWrite);
        9: #Done := "FRK_PersistValidate"(ExpectedKey := "FRK_PersistRuntime".KeyCrc[9], Bytes := "FRK_PersistBuffers".D009Data, Check := "FRK_PersistRuntime".CheckWrite);
        10: #Done := "FRK_PersistValidate"(ExpectedKey := "FRK_PersistRuntime".KeyCrc[10], Bytes := "FRK_PersistBuffers".D010Data, Check := "FRK_PersistRuntime".CheckWrite);
        11: #Done := "FRK_PersistValidate"(ExpectedKey := "FRK_PersistRuntime".KeyCrc[11], Bytes := "FRK_PersistBuffers".D011Data, Check := "FRK_PersistRuntime".CheckWrite);
        12: #Done := "FRK_PersistValidate"(ExpectedKey := "FRK_PersistRuntime".KeyCrc[12], Bytes := "FRK_PersistBuffers".D012Data, Check := "FRK_PersistRuntime".CheckWrite);
        13: #Done := "FRK_PersistValidate"(ExpectedKey := "FRK_PersistRuntime".KeyCrc[13], Bytes := "FRK_PersistBuffers".D013Data, Check := "FRK_PersistRuntime".CheckWrite);
        14: #Done := "FRK_PersistValidate"(ExpectedKey := "FRK_PersistRuntime".KeyCrc[14], Bytes := "FRK_PersistBuffers".D014Data, Check := "FRK_PersistRuntime".CheckWrite);
        15: #Done := "FRK_PersistValidate"(ExpectedKey := "FRK_PersistRuntime".KeyCrc[15], Bytes := "FRK_PersistBuffers".D015Data, Check := "FRK_PersistRuntime".CheckWrite);
        16: #Done := "FRK_PersistValidate"(ExpectedKey := "FRK_PersistRuntime".KeyCrc[16], Bytes := "FRK_PersistBuffers".D016Data, Check := "FRK_PersistRuntime".CheckWrite);
        17: #Done := "FRK_PersistValidate"(ExpectedKey := "FRK_PersistRuntime".KeyCrc[17], Bytes := "FRK_PersistBuffers".D017Data, Check := "FRK_PersistRuntime".CheckWrite);
        18: #Done := "FRK_PersistValidate"(ExpectedKey := "FRK_PersistRuntime".KeyCrc[18], Bytes := "FRK_PersistBuffers".D018Data, Check := "FRK_PersistRuntime".CheckWrite);
        ELSE RETURN;
    END_CASE;
    #FRK_PersistCheckWrite := #Done;
END_FUNCTION
FUNCTION "FRK_PersistInspectSlot" : Void
{ S7_Optimized_Access := 'TRUE' }
VERSION : 0.1
VAR_TEMP
    Done : Bool;
END_VAR
BEGIN
    #Done := FALSE;
    CASE "FRK_PersistRuntime".Slot OF
        1: "FRK_PersistInspect"(BytesA := "FRK_PersistBuffers".D001A, BytesB := "FRK_PersistBuffers".D001B, Payload := "FRK_PersistBuffers".D001Data);
        2: "FRK_PersistInspect"(BytesA := "FRK_PersistBuffers".D002A, BytesB := "FRK_PersistBuffers".D002B, Payload := "FRK_PersistBuffers".D002Data);
        3: "FRK_PersistInspect"(BytesA := "FRK_PersistBuffers".D003A, BytesB := "FRK_PersistBuffers".D003B, Payload := "FRK_PersistBuffers".D003Data);
        4: "FRK_PersistInspect"(BytesA := "FRK_PersistBuffers".D004A, BytesB := "FRK_PersistBuffers".D004B, Payload := "FRK_PersistBuffers".D004Data);
        5: "FRK_PersistInspect"(BytesA := "FRK_PersistBuffers".D005A, BytesB := "FRK_PersistBuffers".D005B, Payload := "FRK_PersistBuffers".D005Data);
        6: "FRK_PersistInspect"(BytesA := "FRK_PersistBuffers".D006A, BytesB := "FRK_PersistBuffers".D006B, Payload := "FRK_PersistBuffers".D006Data);
        7: "FRK_PersistInspect"(BytesA := "FRK_PersistBuffers".D007A, BytesB := "FRK_PersistBuffers".D007B, Payload := "FRK_PersistBuffers".D007Data);
        8: "FRK_PersistInspect"(BytesA := "FRK_PersistBuffers".D008A, BytesB := "FRK_PersistBuffers".D008B, Payload := "FRK_PersistBuffers".D008Data);
        9: "FRK_PersistInspect"(BytesA := "FRK_PersistBuffers".D009A, BytesB := "FRK_PersistBuffers".D009B, Payload := "FRK_PersistBuffers".D009Data);
        10: "FRK_PersistInspect"(BytesA := "FRK_PersistBuffers".D010A, BytesB := "FRK_PersistBuffers".D010B, Payload := "FRK_PersistBuffers".D010Data);
        11: "FRK_PersistInspect"(BytesA := "FRK_PersistBuffers".D011A, BytesB := "FRK_PersistBuffers".D011B, Payload := "FRK_PersistBuffers".D011Data);
        12: "FRK_PersistInspect"(BytesA := "FRK_PersistBuffers".D012A, BytesB := "FRK_PersistBuffers".D012B, Payload := "FRK_PersistBuffers".D012Data);
        13: "FRK_PersistInspect"(BytesA := "FRK_PersistBuffers".D013A, BytesB := "FRK_PersistBuffers".D013B, Payload := "FRK_PersistBuffers".D013Data);
        14: "FRK_PersistInspect"(BytesA := "FRK_PersistBuffers".D014A, BytesB := "FRK_PersistBuffers".D014B, Payload := "FRK_PersistBuffers".D014Data);
        15: "FRK_PersistInspect"(BytesA := "FRK_PersistBuffers".D015A, BytesB := "FRK_PersistBuffers".D015B, Payload := "FRK_PersistBuffers".D015Data);
        16: "FRK_PersistInspect"(BytesA := "FRK_PersistBuffers".D016A, BytesB := "FRK_PersistBuffers".D016B, Payload := "FRK_PersistBuffers".D016Data);
        17: "FRK_PersistInspect"(BytesA := "FRK_PersistBuffers".D017A, BytesB := "FRK_PersistBuffers".D017B, Payload := "FRK_PersistBuffers".D017Data);
        18: "FRK_PersistInspect"(BytesA := "FRK_PersistBuffers".D018A, BytesB := "FRK_PersistBuffers".D018B, Payload := "FRK_PersistBuffers".D018Data);
        ELSE RETURN;
    END_CASE;
END_FUNCTION
FUNCTION "FRK_PersistEnter" : Void
{ S7_Optimized_Access := 'TRUE' }
VERSION : 0.1
VAR_INPUT
    Startup : Bool;
END_VAR
VAR_TEMP
    Index : Int;
END_VAR
BEGIN
    IF #Startup THEN
        "FRK_PersistRuntime".Active := 0; "FRK_PersistRuntime".Stage := 0;
        "FRK_PersistRuntime".HadWrite := TRUE; "FRK_PersistRuntime".LastWriteMs := "FRK_Clock".NowMs; "FRK_PersistRuntime".LastScan := "FRK_PersistRuntime".Scan;
        FOR #Index := 1 TO 4 DO "FRK_PersistRuntime".Queue[#Index].State := 0; END_FOR;
        "FRK_PersistRuntime".Leased[1] := FALSE;
        "FRK_PersistRuntime".Capacity[1] := 13226;
        "FRK_PersistRuntime".KeyCrc[1] := "FRK_PersistKeyCrc"(Key := 'StationA.station');
        IF "FRK_PersistAnchors".SelectedB[1] THEN "FRK_PersistRuntime".Anchor[1] := "FRK_PersistAnchors".RowsB[1]; ELSE "FRK_PersistRuntime".Anchor[1] := "FRK_PersistAnchors".RowsA[1]; END_IF;
        IF NOT "FRK_PersistAnchors".Commissioned[1] AND "FRK_PersistRuntime".Anchor[1].SchemaVersion = 0 AND "FRK_PersistRuntime".Anchor[1].Generation = 0 AND "FRK_PersistRuntime".Anchor[1].KeyCrc = DWORD#0 AND "FRK_PersistRuntime".Anchor[1].DocumentCrc = DWORD#0 AND "FRK_PersistRuntime".Anchor[1].Checksum = DWORD#0 THEN
            "FRK_PersistRepair"(Slot := 1);
        END_IF;
        "FRK_PersistRuntime".Leased[2] := FALSE;
        "FRK_PersistRuntime".Capacity[2] := 12302;
        "FRK_PersistRuntime".KeyCrc[2] := "FRK_PersistKeyCrc"(Key := 'StationA.model.MODEL_A');
        IF "FRK_PersistAnchors".SelectedB[2] THEN "FRK_PersistRuntime".Anchor[2] := "FRK_PersistAnchors".RowsB[2]; ELSE "FRK_PersistRuntime".Anchor[2] := "FRK_PersistAnchors".RowsA[2]; END_IF;
        IF NOT "FRK_PersistAnchors".Commissioned[2] AND "FRK_PersistRuntime".Anchor[2].SchemaVersion = 0 AND "FRK_PersistRuntime".Anchor[2].Generation = 0 AND "FRK_PersistRuntime".Anchor[2].KeyCrc = DWORD#0 AND "FRK_PersistRuntime".Anchor[2].DocumentCrc = DWORD#0 AND "FRK_PersistRuntime".Anchor[2].Checksum = DWORD#0 THEN
            "FRK_PersistRepair"(Slot := 2);
        END_IF;
        "FRK_PersistRuntime".Leased[3] := FALSE;
        "FRK_PersistRuntime".Capacity[3] := 12302;
        "FRK_PersistRuntime".KeyCrc[3] := "FRK_PersistKeyCrc"(Key := 'StationA.model.MODEL_B');
        IF "FRK_PersistAnchors".SelectedB[3] THEN "FRK_PersistRuntime".Anchor[3] := "FRK_PersistAnchors".RowsB[3]; ELSE "FRK_PersistRuntime".Anchor[3] := "FRK_PersistAnchors".RowsA[3]; END_IF;
        IF NOT "FRK_PersistAnchors".Commissioned[3] AND "FRK_PersistRuntime".Anchor[3].SchemaVersion = 0 AND "FRK_PersistRuntime".Anchor[3].Generation = 0 AND "FRK_PersistRuntime".Anchor[3].KeyCrc = DWORD#0 AND "FRK_PersistRuntime".Anchor[3].DocumentCrc = DWORD#0 AND "FRK_PersistRuntime".Anchor[3].Checksum = DWORD#0 THEN
            "FRK_PersistRepair"(Slot := 3);
        END_IF;
        "FRK_PersistRuntime".Leased[4] := FALSE;
        "FRK_PersistRuntime".Capacity[4] := 390;
        "FRK_PersistRuntime".KeyCrc[4] := "FRK_PersistKeyCrc"(Key := 'StationA.policy');
        IF "FRK_PersistAnchors".SelectedB[4] THEN "FRK_PersistRuntime".Anchor[4] := "FRK_PersistAnchors".RowsB[4]; ELSE "FRK_PersistRuntime".Anchor[4] := "FRK_PersistAnchors".RowsA[4]; END_IF;
        IF NOT "FRK_PersistAnchors".Commissioned[4] AND "FRK_PersistRuntime".Anchor[4].SchemaVersion = 0 AND "FRK_PersistRuntime".Anchor[4].Generation = 0 AND "FRK_PersistRuntime".Anchor[4].KeyCrc = DWORD#0 AND "FRK_PersistRuntime".Anchor[4].DocumentCrc = DWORD#0 AND "FRK_PersistRuntime".Anchor[4].Checksum = DWORD#0 THEN
            "FRK_PersistRepair"(Slot := 4);
        END_IF;
        "FRK_PersistRuntime".Leased[5] := FALSE;
        "FRK_PersistRuntime".Capacity[5] := 11186;
        "FRK_PersistRuntime".KeyCrc[5] := "FRK_PersistKeyCrc"(Key := 'StationA.set1');
        IF "FRK_PersistAnchors".SelectedB[5] THEN "FRK_PersistRuntime".Anchor[5] := "FRK_PersistAnchors".RowsB[5]; ELSE "FRK_PersistRuntime".Anchor[5] := "FRK_PersistAnchors".RowsA[5]; END_IF;
        IF NOT "FRK_PersistAnchors".Commissioned[5] AND "FRK_PersistRuntime".Anchor[5].SchemaVersion = 0 AND "FRK_PersistRuntime".Anchor[5].Generation = 0 AND "FRK_PersistRuntime".Anchor[5].KeyCrc = DWORD#0 AND "FRK_PersistRuntime".Anchor[5].DocumentCrc = DWORD#0 AND "FRK_PersistRuntime".Anchor[5].Checksum = DWORD#0 THEN
            "FRK_PersistRepair"(Slot := 5);
        END_IF;
        "FRK_PersistRuntime".Leased[6] := FALSE;
        "FRK_PersistRuntime".Capacity[6] := 11186;
        "FRK_PersistRuntime".KeyCrc[6] := "FRK_PersistKeyCrc"(Key := 'StationA.set2');
        IF "FRK_PersistAnchors".SelectedB[6] THEN "FRK_PersistRuntime".Anchor[6] := "FRK_PersistAnchors".RowsB[6]; ELSE "FRK_PersistRuntime".Anchor[6] := "FRK_PersistAnchors".RowsA[6]; END_IF;
        IF NOT "FRK_PersistAnchors".Commissioned[6] AND "FRK_PersistRuntime".Anchor[6].SchemaVersion = 0 AND "FRK_PersistRuntime".Anchor[6].Generation = 0 AND "FRK_PersistRuntime".Anchor[6].KeyCrc = DWORD#0 AND "FRK_PersistRuntime".Anchor[6].DocumentCrc = DWORD#0 AND "FRK_PersistRuntime".Anchor[6].Checksum = DWORD#0 THEN
            "FRK_PersistRepair"(Slot := 6);
        END_IF;
        "FRK_PersistRuntime".Leased[7] := FALSE;
        "FRK_PersistRuntime".Capacity[7] := 11186;
        "FRK_PersistRuntime".KeyCrc[7] := "FRK_PersistKeyCrc"(Key := 'StationA.set3');
        IF "FRK_PersistAnchors".SelectedB[7] THEN "FRK_PersistRuntime".Anchor[7] := "FRK_PersistAnchors".RowsB[7]; ELSE "FRK_PersistRuntime".Anchor[7] := "FRK_PersistAnchors".RowsA[7]; END_IF;
        IF NOT "FRK_PersistAnchors".Commissioned[7] AND "FRK_PersistRuntime".Anchor[7].SchemaVersion = 0 AND "FRK_PersistRuntime".Anchor[7].Generation = 0 AND "FRK_PersistRuntime".Anchor[7].KeyCrc = DWORD#0 AND "FRK_PersistRuntime".Anchor[7].DocumentCrc = DWORD#0 AND "FRK_PersistRuntime".Anchor[7].Checksum = DWORD#0 THEN
            "FRK_PersistRepair"(Slot := 7);
        END_IF;
        "FRK_PersistRuntime".Leased[8] := FALSE;
        "FRK_PersistRuntime".Capacity[8] := 11186;
        "FRK_PersistRuntime".KeyCrc[8] := "FRK_PersistKeyCrc"(Key := 'StationA.set4');
        IF "FRK_PersistAnchors".SelectedB[8] THEN "FRK_PersistRuntime".Anchor[8] := "FRK_PersistAnchors".RowsB[8]; ELSE "FRK_PersistRuntime".Anchor[8] := "FRK_PersistAnchors".RowsA[8]; END_IF;
        IF NOT "FRK_PersistAnchors".Commissioned[8] AND "FRK_PersistRuntime".Anchor[8].SchemaVersion = 0 AND "FRK_PersistRuntime".Anchor[8].Generation = 0 AND "FRK_PersistRuntime".Anchor[8].KeyCrc = DWORD#0 AND "FRK_PersistRuntime".Anchor[8].DocumentCrc = DWORD#0 AND "FRK_PersistRuntime".Anchor[8].Checksum = DWORD#0 THEN
            "FRK_PersistRepair"(Slot := 8);
        END_IF;
        "FRK_PersistRuntime".Leased[9] := FALSE;
        "FRK_PersistRuntime".Capacity[9] := 13226;
        "FRK_PersistRuntime".KeyCrc[9] := "FRK_PersistKeyCrc"(Key := 'StationB.station');
        IF "FRK_PersistAnchors".SelectedB[9] THEN "FRK_PersistRuntime".Anchor[9] := "FRK_PersistAnchors".RowsB[9]; ELSE "FRK_PersistRuntime".Anchor[9] := "FRK_PersistAnchors".RowsA[9]; END_IF;
        IF NOT "FRK_PersistAnchors".Commissioned[9] AND "FRK_PersistRuntime".Anchor[9].SchemaVersion = 0 AND "FRK_PersistRuntime".Anchor[9].Generation = 0 AND "FRK_PersistRuntime".Anchor[9].KeyCrc = DWORD#0 AND "FRK_PersistRuntime".Anchor[9].DocumentCrc = DWORD#0 AND "FRK_PersistRuntime".Anchor[9].Checksum = DWORD#0 THEN
            "FRK_PersistRepair"(Slot := 9);
        END_IF;
        "FRK_PersistRuntime".Leased[10] := FALSE;
        "FRK_PersistRuntime".Capacity[10] := 12302;
        "FRK_PersistRuntime".KeyCrc[10] := "FRK_PersistKeyCrc"(Key := 'StationB.model.MODEL_A');
        IF "FRK_PersistAnchors".SelectedB[10] THEN "FRK_PersistRuntime".Anchor[10] := "FRK_PersistAnchors".RowsB[10]; ELSE "FRK_PersistRuntime".Anchor[10] := "FRK_PersistAnchors".RowsA[10]; END_IF;
        IF NOT "FRK_PersistAnchors".Commissioned[10] AND "FRK_PersistRuntime".Anchor[10].SchemaVersion = 0 AND "FRK_PersistRuntime".Anchor[10].Generation = 0 AND "FRK_PersistRuntime".Anchor[10].KeyCrc = DWORD#0 AND "FRK_PersistRuntime".Anchor[10].DocumentCrc = DWORD#0 AND "FRK_PersistRuntime".Anchor[10].Checksum = DWORD#0 THEN
            "FRK_PersistRepair"(Slot := 10);
        END_IF;
        "FRK_PersistRuntime".Leased[11] := FALSE;
        "FRK_PersistRuntime".Capacity[11] := 12302;
        "FRK_PersistRuntime".KeyCrc[11] := "FRK_PersistKeyCrc"(Key := 'StationB.model.MODEL_B');
        IF "FRK_PersistAnchors".SelectedB[11] THEN "FRK_PersistRuntime".Anchor[11] := "FRK_PersistAnchors".RowsB[11]; ELSE "FRK_PersistRuntime".Anchor[11] := "FRK_PersistAnchors".RowsA[11]; END_IF;
        IF NOT "FRK_PersistAnchors".Commissioned[11] AND "FRK_PersistRuntime".Anchor[11].SchemaVersion = 0 AND "FRK_PersistRuntime".Anchor[11].Generation = 0 AND "FRK_PersistRuntime".Anchor[11].KeyCrc = DWORD#0 AND "FRK_PersistRuntime".Anchor[11].DocumentCrc = DWORD#0 AND "FRK_PersistRuntime".Anchor[11].Checksum = DWORD#0 THEN
            "FRK_PersistRepair"(Slot := 11);
        END_IF;
        "FRK_PersistRuntime".Leased[12] := FALSE;
        "FRK_PersistRuntime".Capacity[12] := 390;
        "FRK_PersistRuntime".KeyCrc[12] := "FRK_PersistKeyCrc"(Key := 'StationB.policy');
        IF "FRK_PersistAnchors".SelectedB[12] THEN "FRK_PersistRuntime".Anchor[12] := "FRK_PersistAnchors".RowsB[12]; ELSE "FRK_PersistRuntime".Anchor[12] := "FRK_PersistAnchors".RowsA[12]; END_IF;
        IF NOT "FRK_PersistAnchors".Commissioned[12] AND "FRK_PersistRuntime".Anchor[12].SchemaVersion = 0 AND "FRK_PersistRuntime".Anchor[12].Generation = 0 AND "FRK_PersistRuntime".Anchor[12].KeyCrc = DWORD#0 AND "FRK_PersistRuntime".Anchor[12].DocumentCrc = DWORD#0 AND "FRK_PersistRuntime".Anchor[12].Checksum = DWORD#0 THEN
            "FRK_PersistRepair"(Slot := 12);
        END_IF;
        "FRK_PersistRuntime".Leased[13] := FALSE;
        "FRK_PersistRuntime".Capacity[13] := 11186;
        "FRK_PersistRuntime".KeyCrc[13] := "FRK_PersistKeyCrc"(Key := 'StationB.set1');
        IF "FRK_PersistAnchors".SelectedB[13] THEN "FRK_PersistRuntime".Anchor[13] := "FRK_PersistAnchors".RowsB[13]; ELSE "FRK_PersistRuntime".Anchor[13] := "FRK_PersistAnchors".RowsA[13]; END_IF;
        IF NOT "FRK_PersistAnchors".Commissioned[13] AND "FRK_PersistRuntime".Anchor[13].SchemaVersion = 0 AND "FRK_PersistRuntime".Anchor[13].Generation = 0 AND "FRK_PersistRuntime".Anchor[13].KeyCrc = DWORD#0 AND "FRK_PersistRuntime".Anchor[13].DocumentCrc = DWORD#0 AND "FRK_PersistRuntime".Anchor[13].Checksum = DWORD#0 THEN
            "FRK_PersistRepair"(Slot := 13);
        END_IF;
        "FRK_PersistRuntime".Leased[14] := FALSE;
        "FRK_PersistRuntime".Capacity[14] := 11186;
        "FRK_PersistRuntime".KeyCrc[14] := "FRK_PersistKeyCrc"(Key := 'StationB.set2');
        IF "FRK_PersistAnchors".SelectedB[14] THEN "FRK_PersistRuntime".Anchor[14] := "FRK_PersistAnchors".RowsB[14]; ELSE "FRK_PersistRuntime".Anchor[14] := "FRK_PersistAnchors".RowsA[14]; END_IF;
        IF NOT "FRK_PersistAnchors".Commissioned[14] AND "FRK_PersistRuntime".Anchor[14].SchemaVersion = 0 AND "FRK_PersistRuntime".Anchor[14].Generation = 0 AND "FRK_PersistRuntime".Anchor[14].KeyCrc = DWORD#0 AND "FRK_PersistRuntime".Anchor[14].DocumentCrc = DWORD#0 AND "FRK_PersistRuntime".Anchor[14].Checksum = DWORD#0 THEN
            "FRK_PersistRepair"(Slot := 14);
        END_IF;
        "FRK_PersistRuntime".Leased[15] := FALSE;
        "FRK_PersistRuntime".Capacity[15] := 11186;
        "FRK_PersistRuntime".KeyCrc[15] := "FRK_PersistKeyCrc"(Key := 'StationB.set3');
        IF "FRK_PersistAnchors".SelectedB[15] THEN "FRK_PersistRuntime".Anchor[15] := "FRK_PersistAnchors".RowsB[15]; ELSE "FRK_PersistRuntime".Anchor[15] := "FRK_PersistAnchors".RowsA[15]; END_IF;
        IF NOT "FRK_PersistAnchors".Commissioned[15] AND "FRK_PersistRuntime".Anchor[15].SchemaVersion = 0 AND "FRK_PersistRuntime".Anchor[15].Generation = 0 AND "FRK_PersistRuntime".Anchor[15].KeyCrc = DWORD#0 AND "FRK_PersistRuntime".Anchor[15].DocumentCrc = DWORD#0 AND "FRK_PersistRuntime".Anchor[15].Checksum = DWORD#0 THEN
            "FRK_PersistRepair"(Slot := 15);
        END_IF;
        "FRK_PersistRuntime".Leased[16] := FALSE;
        "FRK_PersistRuntime".Capacity[16] := 11186;
        "FRK_PersistRuntime".KeyCrc[16] := "FRK_PersistKeyCrc"(Key := 'StationB.set4');
        IF "FRK_PersistAnchors".SelectedB[16] THEN "FRK_PersistRuntime".Anchor[16] := "FRK_PersistAnchors".RowsB[16]; ELSE "FRK_PersistRuntime".Anchor[16] := "FRK_PersistAnchors".RowsA[16]; END_IF;
        IF NOT "FRK_PersistAnchors".Commissioned[16] AND "FRK_PersistRuntime".Anchor[16].SchemaVersion = 0 AND "FRK_PersistRuntime".Anchor[16].Generation = 0 AND "FRK_PersistRuntime".Anchor[16].KeyCrc = DWORD#0 AND "FRK_PersistRuntime".Anchor[16].DocumentCrc = DWORD#0 AND "FRK_PersistRuntime".Anchor[16].Checksum = DWORD#0 THEN
            "FRK_PersistRepair"(Slot := 16);
        END_IF;
        "FRK_PersistRuntime".Leased[17] := FALSE;
        "FRK_PersistRuntime".Capacity[17] := 8704;
        "FRK_PersistRuntime".KeyCrc[17] := "FRK_PersistKeyCrc"(Key := 'users');
        IF "FRK_PersistAnchors".SelectedB[17] THEN "FRK_PersistRuntime".Anchor[17] := "FRK_PersistAnchors".RowsB[17]; ELSE "FRK_PersistRuntime".Anchor[17] := "FRK_PersistAnchors".RowsA[17]; END_IF;
        IF NOT "FRK_PersistAnchors".Commissioned[17] AND "FRK_PersistRuntime".Anchor[17].SchemaVersion = 0 AND "FRK_PersistRuntime".Anchor[17].Generation = 0 AND "FRK_PersistRuntime".Anchor[17].KeyCrc = DWORD#0 AND "FRK_PersistRuntime".Anchor[17].DocumentCrc = DWORD#0 AND "FRK_PersistRuntime".Anchor[17].Checksum = DWORD#0 THEN
            "FRK_PersistRepair"(Slot := 17);
        END_IF;
        "FRK_PersistRuntime".Leased[18] := FALSE;
        "FRK_PersistRuntime".Capacity[18] := 8732;
        "FRK_PersistRuntime".KeyCrc[18] := "FRK_PersistKeyCrc"(Key := 'line.76378c768007b72db223c2939faaa0e1e06be912b0a3ff238e89cbb24ff9effd');
        IF "FRK_PersistAnchors".SelectedB[18] THEN "FRK_PersistRuntime".Anchor[18] := "FRK_PersistAnchors".RowsB[18]; ELSE "FRK_PersistRuntime".Anchor[18] := "FRK_PersistAnchors".RowsA[18]; END_IF;
        IF NOT "FRK_PersistAnchors".Commissioned[18] AND "FRK_PersistRuntime".Anchor[18].SchemaVersion = 0 AND "FRK_PersistRuntime".Anchor[18].Generation = 0 AND "FRK_PersistRuntime".Anchor[18].KeyCrc = DWORD#0 AND "FRK_PersistRuntime".Anchor[18].DocumentCrc = DWORD#0 AND "FRK_PersistRuntime".Anchor[18].Checksum = DWORD#0 THEN
            "FRK_PersistRepair"(Slot := 18);
        END_IF;
    END_IF;
    "FRK_PersistRuntime".Scan := "FRK_PersistRuntime".Scan + 1;
END_FUNCTION
FUNCTION "FRK_PersistTick" : Void
{ S7_Optimized_Access := 'TRUE' }
VERSION : 0.1
VAR_TEMP
    Pick : Int;
    Index : Int;
    Slot : Int;
    Operation : Int;
    Done : Bool;
    Check : "FRK_PersistCheck";
END_VAR
BEGIN
    IF "FRK_PersistRuntime".LastScan = "FRK_PersistRuntime".Scan THEN RETURN; END_IF;
    "FRK_PersistRuntime".LastScan := "FRK_PersistRuntime".Scan;
    IF "FRK_PersistRuntime".Active = 0 THEN
        #Pick := 0;
        FOR #Index := 1 TO 4 DO
            IF "FRK_PersistRuntime".Queue[#Index].State = 1 THEN
                IF #Pick = 0 THEN #Pick := #Index; ELSIF "FRK_PersistRuntime".Queue[#Index].Ticket < "FRK_PersistRuntime".Queue[#Pick].Ticket THEN #Pick := #Index; END_IF;
            END_IF;
        END_FOR;
        IF #Pick = 0 THEN RETURN; END_IF;
        "FRK_PersistRuntime".Active := #Pick;
        "FRK_PersistRuntime".Slot := "FRK_PersistRuntime".Queue[#Pick].Slot;
        "FRK_PersistRuntime".Queue[#Pick].State := 2;
        "FRK_PersistRuntime".Result := "FRK_PersistRuntime".EmptyResult;
        "FRK_PersistRuntime".Stage := 1; "FRK_PersistRuntime".NativeReq := TRUE;
        "FRK_PersistRuntime".CheckA.Cursor := -1; "FRK_PersistRuntime".CheckB.Cursor := -1;
    END_IF;
    IF "FRK_PersistRuntime".Unavailable THEN
        "FRK_PersistRuntime".Result.ErrorId := UDINT#32963;
        "FRK_PersistFinish"(); RETURN;
    END_IF;
    CASE "FRK_PersistRuntime".Stage OF
        1, 2, 8, 9:
            #Operation := "FRK_PersistRuntime".Stage;
            IF #Operation = 8 THEN #Operation := "FRK_PersistRuntime".Chosen + 2; ELSIF #Operation = 9 THEN #Operation := "FRK_PersistRuntime".Chosen; END_IF;
            "FRK_PersistIo"(Operation := #Operation);
            "FRK_PersistRuntime".NativeReq := FALSE;
            IF "FRK_PersistRuntime".NativeBusy THEN RETURN; END_IF;
            IF "FRK_PersistRuntime".NativeResult <> 0 THEN
                "FRK_PersistRuntime".Result.ErrorId := WORD_TO_UDINT(INT_TO_WORD("FRK_PersistRuntime".NativeResult));
                "FRK_PersistFinish"(); RETURN;
            END_IF;
            CASE "FRK_PersistRuntime".Stage OF
                1: "FRK_PersistRuntime".Stage := 2;
                2: "FRK_PersistRuntime".Stage := 3;
                8: "FRK_PersistRuntime".Stage := 9;
                9: "FRK_PersistRuntime".Stage := 10; IF "FRK_PersistRuntime".Chosen = 1 THEN "FRK_PersistRuntime".CheckA.Cursor := -1; ELSE "FRK_PersistRuntime".CheckB.Cursor := -1; END_IF;
                ELSE RETURN;
            END_CASE;
            "FRK_PersistRuntime".NativeReq := TRUE;
        3: IF "FRK_PersistCheckA"() THEN "FRK_PersistRuntime".Stage := 4; END_IF;
        4: IF "FRK_PersistCheckB"() THEN "FRK_PersistRuntime".Stage := 5; END_IF;
        5: "FRK_PersistInspectSlot"();
        6:
            IF "FRK_PersistCheckWrite"() THEN
                CASE "FRK_PersistRuntime".Slot OF
                    1: "FRK_PersistPutNumber"(Bytes := "FRK_PersistBuffers".D001Data, Offset := 20, Value := "FRK_PersistRuntime".CheckWrite.Crc);
                    2: "FRK_PersistPutNumber"(Bytes := "FRK_PersistBuffers".D002Data, Offset := 20, Value := "FRK_PersistRuntime".CheckWrite.Crc);
                    3: "FRK_PersistPutNumber"(Bytes := "FRK_PersistBuffers".D003Data, Offset := 20, Value := "FRK_PersistRuntime".CheckWrite.Crc);
                    4: "FRK_PersistPutNumber"(Bytes := "FRK_PersistBuffers".D004Data, Offset := 20, Value := "FRK_PersistRuntime".CheckWrite.Crc);
                    5: "FRK_PersistPutNumber"(Bytes := "FRK_PersistBuffers".D005Data, Offset := 20, Value := "FRK_PersistRuntime".CheckWrite.Crc);
                    6: "FRK_PersistPutNumber"(Bytes := "FRK_PersistBuffers".D006Data, Offset := 20, Value := "FRK_PersistRuntime".CheckWrite.Crc);
                    7: "FRK_PersistPutNumber"(Bytes := "FRK_PersistBuffers".D007Data, Offset := 20, Value := "FRK_PersistRuntime".CheckWrite.Crc);
                    8: "FRK_PersistPutNumber"(Bytes := "FRK_PersistBuffers".D008Data, Offset := 20, Value := "FRK_PersistRuntime".CheckWrite.Crc);
                    9: "FRK_PersistPutNumber"(Bytes := "FRK_PersistBuffers".D009Data, Offset := 20, Value := "FRK_PersistRuntime".CheckWrite.Crc);
                    10: "FRK_PersistPutNumber"(Bytes := "FRK_PersistBuffers".D010Data, Offset := 20, Value := "FRK_PersistRuntime".CheckWrite.Crc);
                    11: "FRK_PersistPutNumber"(Bytes := "FRK_PersistBuffers".D011Data, Offset := 20, Value := "FRK_PersistRuntime".CheckWrite.Crc);
                    12: "FRK_PersistPutNumber"(Bytes := "FRK_PersistBuffers".D012Data, Offset := 20, Value := "FRK_PersistRuntime".CheckWrite.Crc);
                    13: "FRK_PersistPutNumber"(Bytes := "FRK_PersistBuffers".D013Data, Offset := 20, Value := "FRK_PersistRuntime".CheckWrite.Crc);
                    14: "FRK_PersistPutNumber"(Bytes := "FRK_PersistBuffers".D014Data, Offset := 20, Value := "FRK_PersistRuntime".CheckWrite.Crc);
                    15: "FRK_PersistPutNumber"(Bytes := "FRK_PersistBuffers".D015Data, Offset := 20, Value := "FRK_PersistRuntime".CheckWrite.Crc);
                    16: "FRK_PersistPutNumber"(Bytes := "FRK_PersistBuffers".D016Data, Offset := 20, Value := "FRK_PersistRuntime".CheckWrite.Crc);
                    17: "FRK_PersistPutNumber"(Bytes := "FRK_PersistBuffers".D017Data, Offset := 20, Value := "FRK_PersistRuntime".CheckWrite.Crc);
                    18: "FRK_PersistPutNumber"(Bytes := "FRK_PersistBuffers".D018Data, Offset := 20, Value := "FRK_PersistRuntime".CheckWrite.Crc);
                    ELSE RETURN;
                END_CASE;
                "FRK_PersistRuntime".Stage := 7;
            END_IF;
        7:
            IF NOT "FRK_PersistRuntime".HadWrite OR "FRK_Elapsed"(OldMs := "FRK_PersistRuntime".LastWriteMs, NewMs := "FRK_Clock".NowMs) >= 1000 THEN
                "FRK_PersistRuntime".HadWrite := TRUE; "FRK_PersistRuntime".LastWriteMs := "FRK_Clock".NowMs;
                "FRK_PersistRuntime".Stage := 8; "FRK_PersistRuntime".NativeReq := TRUE;
            END_IF;
        10:
            IF "FRK_PersistRuntime".Chosen = 1 THEN #Done := "FRK_PersistCheckA"(); #Check := "FRK_PersistRuntime".CheckA;
            ELSE #Done := "FRK_PersistCheckB"(); #Check := "FRK_PersistRuntime".CheckB; END_IF;
            IF #Done THEN
                IF #Check.Valid AND #Check.Generation = "FRK_PersistRuntime".Generation AND #Check.Crc = "FRK_PersistRuntime".CheckWrite.Crc THEN
                    #Slot := "FRK_PersistRuntime".Slot;
                    "FRK_PersistRuntime".Anchor[#Slot].Generation := #Check.Generation;
                    "FRK_PersistRuntime".Anchor[#Slot].DocumentCrc := #Check.Crc;
                    "FRK_PersistRuntime".Anchor[#Slot].Checksum := "FRK_PersistAnchorCrc"(Image := "FRK_PersistRuntime".Anchor[#Slot]);
                    "FRK_PersistCommitAnchor"(Slot := #Slot);
                    "FRK_PersistRuntime".Result.Ok := TRUE;
                ELSE "FRK_PersistRuntime".Result.ErrorId := 4; END_IF;
                "FRK_PersistFinish"();
            END_IF;
        ELSE
            "FRK_PersistRuntime".Result.ErrorId := 1; "FRK_PersistFinish"();
    END_CASE;
END_FUNCTION
FUNCTION "FRK_PersistPoll" : Bool
{ S7_Optimized_Access := 'TRUE' }
VERSION : 0.1
VAR_INPUT
    Ticket : UDInt;
END_VAR
VAR_IN_OUT
    Result : "ST_PersistResult";
END_VAR
VAR_TEMP
    Index : Int;
END_VAR
BEGIN
    #FRK_PersistPoll := TRUE; #Result := "FRK_PersistRuntime".EmptyResult;
    #Result.ErrorId := 1;
    "FRK_PersistTick"();
    IF #Ticket = 0 THEN RETURN; END_IF;
    FOR #Index := 1 TO 4 DO
        IF "FRK_PersistRuntime".Queue[#Index].State <> 0 AND "FRK_PersistRuntime".Queue[#Index].Ticket = #Ticket THEN
            #FRK_PersistPoll := "FRK_PersistRuntime".Queue[#Index].State = 3;
            IF #FRK_PersistPoll THEN
                #Result := "FRK_PersistRuntime".Queue[#Index].Result;
                "FRK_PersistRuntime".Leased["FRK_PersistRuntime".Queue[#Index].Slot] := FALSE;
                "FRK_PersistRuntime".Queue[#Index].State := 0;
            END_IF;
            RETURN;
        END_IF;
    END_FOR;
END_FUNCTION
FUNCTION "FRK_DocCapture_D001" : Bool
{ S7_Optimized_Access := 'TRUE' }
VERSION : 0.1
VAR_IN_OUT
    Length : DInt;
END_VAR
VAR_TEMP
    Index : Int;
    Stored : Int;
    Position : DInt;
    NativeResult : Int;
    Ok : Bool;
    Targets : Array[1..28] of Int;
    Prior : Int;
    Reserved : Bool;
END_VAR
BEGIN
    #FRK_DocCapture_D001 := FALSE;
    "FRK_PersistImages".D001.SchemaVersion := 1; "FRK_PersistImages".D001.Scope := 'StationA';
    "FRK_PersistImages".D001.Kind := 1;
    "FRK_PersistImages".D001.ModelCode := '';
    "FRK_PersistImages".D001.ActiveModel := "FRK_ConfigStore".ActiveModels[1];
    "FRK_PersistImages".D001.Count := 28;
    #Stored := "FRK_ConfigFind"(Scope := 'StationA', Key := 'siteLabel', ModelCode := '');
    IF #Stored = 0 THEN RETURN; END_IF;
    "FRK_PersistImages".D001.Rows[1] := "FRK_ConfigStore".Rows[#Stored];
    #Stored := "FRK_ConfigFind"(Scope := 'StationA', Key := 'enabled', ModelCode := '');
    IF #Stored = 0 THEN RETURN; END_IF;
    "FRK_PersistImages".D001.Rows[2] := "FRK_ConfigStore".Rows[#Stored];
    #Stored := "FRK_ConfigFind"(Scope := 'StationA', Key := 'ratio', ModelCode := '');
    IF #Stored = 0 THEN RETURN; END_IF;
    "FRK_PersistImages".D001.Rows[3] := "FRK_ConfigStore".Rows[#Stored];
    #Stored := "FRK_ConfigFind"(Scope := 'StationA', Key := 'gain', ModelCode := '');
    IF #Stored = 0 THEN RETURN; END_IF;
    "FRK_PersistImages".D001.Rows[4] := "FRK_ConfigStore".Rows[#Stored];
    #Stored := "FRK_ConfigFind"(Scope := 'StationA', Key := 'grade', ModelCode := '');
    IF #Stored = 0 THEN RETURN; END_IF;
    "FRK_PersistImages".D001.Rows[5] := "FRK_ConfigStore".Rows[#Stored];
    #Stored := "FRK_ConfigFind"(Scope := 'StationA', Key := 'small', ModelCode := '');
    IF #Stored = 0 THEN RETURN; END_IF;
    "FRK_PersistImages".D001.Rows[6] := "FRK_ConfigStore".Rows[#Stored];
    #Stored := "FRK_ConfigFind"(Scope := 'StationA', Key := 'long.kkkkkkkkkkkkkkkkkkkkkkkkkkkkkkkkkkkkkkkkkkkkkkkkkkkkkkkkkkkkkkkkkkkkkkkkkkkkkkkkkkkkkkkkkkkkkkkkkkkkkkkkkkkkkkkkkkkkkkkkkkkkkkkkkkkkkkk', ModelCode := '');
    IF #Stored = 0 THEN RETURN; END_IF;
    "FRK_PersistImages".D001.Rows[7] := "FRK_ConfigStore".Rows[#Stored];
    #Stored := "FRK_ConfigFind"(Scope := 'StationA', Key := 'degradationPercent', ModelCode := '');
    IF #Stored = 0 THEN RETURN; END_IF;
    "FRK_PersistImages".D001.Rows[8] := "FRK_ConfigStore".Rows[#Stored];
    #Stored := "FRK_ConfigFind"(Scope := 'StationA.Satellite', Key := 'siteLabel', ModelCode := '');
    IF #Stored = 0 THEN RETURN; END_IF;
    "FRK_PersistImages".D001.Rows[9] := "FRK_ConfigStore".Rows[#Stored];
    #Stored := "FRK_ConfigFind"(Scope := 'StationA.Satellite', Key := 'enabled', ModelCode := '');
    IF #Stored = 0 THEN RETURN; END_IF;
    "FRK_PersistImages".D001.Rows[10] := "FRK_ConfigStore".Rows[#Stored];
    #Stored := "FRK_ConfigFind"(Scope := 'StationA.Satellite', Key := 'ratio', ModelCode := '');
    IF #Stored = 0 THEN RETURN; END_IF;
    "FRK_PersistImages".D001.Rows[11] := "FRK_ConfigStore".Rows[#Stored];
    #Stored := "FRK_ConfigFind"(Scope := 'StationA.Satellite', Key := 'gain', ModelCode := '');
    IF #Stored = 0 THEN RETURN; END_IF;
    "FRK_PersistImages".D001.Rows[12] := "FRK_ConfigStore".Rows[#Stored];
    #Stored := "FRK_ConfigFind"(Scope := 'StationA.Satellite', Key := 'grade', ModelCode := '');
    IF #Stored = 0 THEN RETURN; END_IF;
    "FRK_PersistImages".D001.Rows[13] := "FRK_ConfigStore".Rows[#Stored];
    #Stored := "FRK_ConfigFind"(Scope := 'StationA.Satellite', Key := 'offset.-1', ModelCode := '');
    IF #Stored = 0 THEN RETURN; END_IF;
    "FRK_PersistImages".D001.Rows[14] := "FRK_ConfigStore".Rows[#Stored];
    #Stored := "FRK_ConfigFind"(Scope := 'StationA.Satellite', Key := 'offset.0', ModelCode := '');
    IF #Stored = 0 THEN RETURN; END_IF;
    "FRK_PersistImages".D001.Rows[15] := "FRK_ConfigStore".Rows[#Stored];
    #Stored := "FRK_ConfigFind"(Scope := 'StationA.Satellite', Key := 'offset.1', ModelCode := '');
    IF #Stored = 0 THEN RETURN; END_IF;
    "FRK_PersistImages".D001.Rows[16] := "FRK_ConfigStore".Rows[#Stored];
    #Stored := "FRK_ConfigFind"(Scope := 'StationA.Satellite', Key := 'long.kkkkkkkkkkkkkkkkkkkkkkkkkkkkkkkkkkkkkkkkkkkkkkkkkkkkkkkkkkkkkkkkkkkkkkkkkkkkkkkkkkkkkkkkkkkkkkkkkkkkkkkkkkkkkkkkkkkkkkkkkkkkkkkkkkkkkkk', ModelCode := '');
    IF #Stored = 0 THEN RETURN; END_IF;
    "FRK_PersistImages".D001.Rows[17] := "FRK_ConfigStore".Rows[#Stored];
    #Stored := "FRK_ConfigFind"(Scope := 'StationA.Satellite', Key := 'small', ModelCode := '');
    IF #Stored = 0 THEN RETURN; END_IF;
    "FRK_PersistImages".D001.Rows[18] := "FRK_ConfigStore".Rows[#Stored];
    #Stored := "FRK_ConfigFind"(Scope := 'StationA.Satellite.Inner', Key := 'siteLabel', ModelCode := '');
    IF #Stored = 0 THEN RETURN; END_IF;
    "FRK_PersistImages".D001.Rows[19] := "FRK_ConfigStore".Rows[#Stored];
    #Stored := "FRK_ConfigFind"(Scope := 'StationA.Satellite.Inner', Key := 'enabled', ModelCode := '');
    IF #Stored = 0 THEN RETURN; END_IF;
    "FRK_PersistImages".D001.Rows[20] := "FRK_ConfigStore".Rows[#Stored];
    #Stored := "FRK_ConfigFind"(Scope := 'StationA.Satellite.Inner', Key := 'ratio', ModelCode := '');
    IF #Stored = 0 THEN RETURN; END_IF;
    "FRK_PersistImages".D001.Rows[21] := "FRK_ConfigStore".Rows[#Stored];
    #Stored := "FRK_ConfigFind"(Scope := 'StationA.Satellite.Inner', Key := 'gain', ModelCode := '');
    IF #Stored = 0 THEN RETURN; END_IF;
    "FRK_PersistImages".D001.Rows[22] := "FRK_ConfigStore".Rows[#Stored];
    #Stored := "FRK_ConfigFind"(Scope := 'StationA.Satellite.Inner', Key := 'grade', ModelCode := '');
    IF #Stored = 0 THEN RETURN; END_IF;
    "FRK_PersistImages".D001.Rows[23] := "FRK_ConfigStore".Rows[#Stored];
    #Stored := "FRK_ConfigFind"(Scope := 'StationA.Satellite.Inner', Key := 'offset.-1', ModelCode := '');
    IF #Stored = 0 THEN RETURN; END_IF;
    "FRK_PersistImages".D001.Rows[24] := "FRK_ConfigStore".Rows[#Stored];
    #Stored := "FRK_ConfigFind"(Scope := 'StationA.Satellite.Inner', Key := 'offset.0', ModelCode := '');
    IF #Stored = 0 THEN RETURN; END_IF;
    "FRK_PersistImages".D001.Rows[25] := "FRK_ConfigStore".Rows[#Stored];
    #Stored := "FRK_ConfigFind"(Scope := 'StationA.Satellite.Inner', Key := 'offset.1', ModelCode := '');
    IF #Stored = 0 THEN RETURN; END_IF;
    "FRK_PersistImages".D001.Rows[26] := "FRK_ConfigStore".Rows[#Stored];
    #Stored := "FRK_ConfigFind"(Scope := 'StationA.Satellite.Inner', Key := 'long.kkkkkkkkkkkkkkkkkkkkkkkkkkkkkkkkkkkkkkkkkkkkkkkkkkkkkkkkkkkkkkkkkkkkkkkkkkkkkkkkkkkkkkkkkkkkkkkkkkkkkkkkkkkkkkkkkkkkkkkkkkkkkkkkkkkkkkk', ModelCode := '');
    IF #Stored = 0 THEN RETURN; END_IF;
    "FRK_PersistImages".D001.Rows[27] := "FRK_ConfigStore".Rows[#Stored];
    #Stored := "FRK_ConfigFind"(Scope := 'StationA.Satellite.Inner', Key := 'small', ModelCode := '');
    IF #Stored = 0 THEN RETURN; END_IF;
    "FRK_PersistImages".D001.Rows[28] := "FRK_ConfigStore".Rows[#Stored];
    FOR #Index := 0 TO 13249 DO "FRK_PersistBuffers".D001Data[#Index] := BYTE#0; END_FOR;
    #Position := 24;
    #NativeResult := Serialize(SRC_VARIABLE := "FRK_PersistImages".D001, DEST_ARRAY => "FRK_PersistBuffers".D001Data, POS := #Position);
    IF #NativeResult <> 0 OR #Position < 24 OR #Position > 13250 THEN RETURN; END_IF;
    #Length := #Position - 24;
    #FRK_DocCapture_D001 := TRUE;
END_FUNCTION
FUNCTION "FRK_DocApply_D001" : Bool
{ S7_Optimized_Access := 'TRUE' }
VERSION : 0.1
VAR_TEMP
    Index : Int;
    Stored : Int;
    Position : DInt;
    NativeResult : Int;
    Ok : Bool;
    Targets : Array[1..28] of Int;
    Prior : Int;
    Reserved : Bool;
END_VAR
BEGIN
    #FRK_DocApply_D001 := FALSE;
    #Position := 24;
    #NativeResult := Deserialize(SRC_ARRAY := "FRK_PersistBuffers".D001Data, DEST_VARIABLE => "FRK_PersistImages".D001, POS := #Position);
    IF #NativeResult <> 0 OR #Position <> 24 + UDINT_TO_DINT("FRK_PersistConsumers".Rows[1].Result.Length) THEN RETURN; END_IF;
    IF "FRK_PersistImages".D001.SchemaVersion <> 1 OR "FRK_PersistImages".D001.Scope <> 'StationA' THEN RETURN; END_IF;
    IF "FRK_PersistImages".D001.Kind <> 1 OR "FRK_PersistImages".D001.ModelCode <> '' OR "FRK_PersistImages".D001.Count <> 28 THEN RETURN; END_IF;
    IF "FRK_PersistImages".D001.ActiveModel <> 'MODEL_A' AND "FRK_PersistImages".D001.ActiveModel <> 'MODEL_B' THEN RETURN; END_IF;
    IF NOT "FRK_PersistImages".D001.Rows[1].Used OR "FRK_PersistImages".D001.Rows[1].SchemaVersion <> 3 OR "FRK_PersistImages".D001.Rows[1].ModelCode <> '' OR "FRK_PersistImages".D001.Rows[1].Record.Scope <> 'StationA' OR "FRK_PersistImages".D001.Rows[1].Record.WriteKey <> 'siteLabel' OR "FRK_PersistImages".D001.Rows[1].Record.Revision <> 1 OR "FRK_PersistImages".D001.Rows[1].Record.Kind <> 1 OR "FRK_PersistImages".D001.Rows[1].Record.ValueType <> 1 THEN RETURN; END_IF;
    #Ok := "FRK_ConfigDecode"(Text := STRING_TO_WSTRING("FRK_PersistImages".D001.Rows[1].Record.ValueText), Storage := 8, Minimum := 0.0, Maximum := 1.0, MaxLength := 80, Value := "FRK_ConfigScratch".Value);
    IF NOT #Ok THEN RETURN; END_IF;
    IF NOT "FRK_PersistImages".D001.Rows[2].Used OR "FRK_PersistImages".D001.Rows[2].SchemaVersion <> 3 OR "FRK_PersistImages".D001.Rows[2].ModelCode <> '' OR "FRK_PersistImages".D001.Rows[2].Record.Scope <> 'StationA' OR "FRK_PersistImages".D001.Rows[2].Record.WriteKey <> 'enabled' OR "FRK_PersistImages".D001.Rows[2].Record.Revision <> 1 OR "FRK_PersistImages".D001.Rows[2].Record.Kind <> 1 OR "FRK_PersistImages".D001.Rows[2].Record.ValueType <> 2 THEN RETURN; END_IF;
    #Ok := "FRK_ConfigDecode"(Text := STRING_TO_WSTRING("FRK_PersistImages".D001.Rows[2].Record.ValueText), Storage := 1, Minimum := 0.0, Maximum := 1.0, MaxLength := 0, Value := "FRK_ConfigScratch".Value);
    IF NOT #Ok THEN RETURN; END_IF;
    IF NOT "FRK_PersistImages".D001.Rows[3].Used OR "FRK_PersistImages".D001.Rows[3].SchemaVersion <> 3 OR "FRK_PersistImages".D001.Rows[3].ModelCode <> '' OR "FRK_PersistImages".D001.Rows[3].Record.Scope <> 'StationA' OR "FRK_PersistImages".D001.Rows[3].Record.WriteKey <> 'ratio' OR "FRK_PersistImages".D001.Rows[3].Record.Revision <> 1 OR "FRK_PersistImages".D001.Rows[3].Record.Kind <> 1 OR "FRK_PersistImages".D001.Rows[3].Record.ValueType <> 0 THEN RETURN; END_IF;
    #Ok := "FRK_ConfigDecode"(Text := STRING_TO_WSTRING("FRK_PersistImages".D001.Rows[3].Record.ValueText), Storage := 6, Minimum := -1000000.0, Maximum := 1000000.0, MaxLength := 0, Value := "FRK_ConfigScratch".Value);
    IF NOT #Ok THEN RETURN; END_IF;
    IF NOT "FRK_PersistImages".D001.Rows[4].Used OR "FRK_PersistImages".D001.Rows[4].SchemaVersion <> 3 OR "FRK_PersistImages".D001.Rows[4].ModelCode <> '' OR "FRK_PersistImages".D001.Rows[4].Record.Scope <> 'StationA' OR "FRK_PersistImages".D001.Rows[4].Record.WriteKey <> 'gain' OR "FRK_PersistImages".D001.Rows[4].Record.Revision <> 1 OR "FRK_PersistImages".D001.Rows[4].Record.Kind <> 1 OR "FRK_PersistImages".D001.Rows[4].Record.ValueType <> 0 THEN RETURN; END_IF;
    #Ok := "FRK_ConfigDecode"(Text := STRING_TO_WSTRING("FRK_PersistImages".D001.Rows[4].Record.ValueText), Storage := 5, Minimum := -1000.0, Maximum := 1000.0, MaxLength := 0, Value := "FRK_ConfigScratch".Value);
    IF NOT #Ok THEN RETURN; END_IF;
    IF NOT "FRK_PersistImages".D001.Rows[5].Used OR "FRK_PersistImages".D001.Rows[5].SchemaVersion <> 3 OR "FRK_PersistImages".D001.Rows[5].ModelCode <> '' OR "FRK_PersistImages".D001.Rows[5].Record.Scope <> 'StationA' OR "FRK_PersistImages".D001.Rows[5].Record.WriteKey <> 'grade' OR "FRK_PersistImages".D001.Rows[5].Record.Revision <> 1 OR "FRK_PersistImages".D001.Rows[5].Record.Kind <> 1 OR "FRK_PersistImages".D001.Rows[5].Record.ValueType <> 0 THEN RETURN; END_IF;
    #Ok := "FRK_ConfigDecode"(Text := STRING_TO_WSTRING("FRK_PersistImages".D001.Rows[5].Record.ValueText), Storage := 3, Minimum := 0.0, Maximum := 6.0, MaxLength := 0, Value := "FRK_ConfigScratch".Value);
    IF NOT #Ok THEN RETURN; END_IF;
    IF NOT "FRK_PersistImages".D001.Rows[6].Used OR "FRK_PersistImages".D001.Rows[6].SchemaVersion <> 3 OR "FRK_PersistImages".D001.Rows[6].ModelCode <> '' OR "FRK_PersistImages".D001.Rows[6].Record.Scope <> 'StationA' OR "FRK_PersistImages".D001.Rows[6].Record.WriteKey <> 'small' OR "FRK_PersistImages".D001.Rows[6].Record.Revision <> 1 OR "FRK_PersistImages".D001.Rows[6].Record.Kind <> 1 OR "FRK_PersistImages".D001.Rows[6].Record.ValueType <> 0 THEN RETURN; END_IF;
    #Ok := "FRK_ConfigDecode"(Text := STRING_TO_WSTRING("FRK_PersistImages".D001.Rows[6].Record.ValueText), Storage := 3, Minimum := 0.0, Maximum := 255.0, MaxLength := 0, Value := "FRK_ConfigScratch".Value);
    IF NOT #Ok THEN RETURN; END_IF;
    IF NOT "FRK_PersistImages".D001.Rows[7].Used OR "FRK_PersistImages".D001.Rows[7].SchemaVersion <> 3 OR "FRK_PersistImages".D001.Rows[7].ModelCode <> '' OR "FRK_PersistImages".D001.Rows[7].Record.Scope <> 'StationA' OR "FRK_PersistImages".D001.Rows[7].Record.WriteKey <> 'long.kkkkkkkkkkkkkkkkkkkkkkkkkkkkkkkkkkkkkkkkkkkkkkkkkkkkkkkkkkkkkkkkkkkkkkkkkkkkkkkkkkkkkkkkkkkkkkkkkkkkkkkkkkkkkkkkkkkkkkkkkkkkkkkkkkkkkkk' OR "FRK_PersistImages".D001.Rows[7].Record.Revision <> 1 OR "FRK_PersistImages".D001.Rows[7].Record.Kind <> 1 OR "FRK_PersistImages".D001.Rows[7].Record.ValueType <> 1 THEN RETURN; END_IF;
    #Ok := "FRK_ConfigDecode"(Text := STRING_TO_WSTRING("FRK_PersistImages".D001.Rows[7].Record.ValueText), Storage := 8, Minimum := 0.0, Maximum := 1.0, MaxLength := 80, Value := "FRK_ConfigScratch".Value);
    IF NOT #Ok THEN RETURN; END_IF;
    IF NOT "FRK_PersistImages".D001.Rows[8].Used OR "FRK_PersistImages".D001.Rows[8].SchemaVersion <> 3 OR "FRK_PersistImages".D001.Rows[8].ModelCode <> '' OR "FRK_PersistImages".D001.Rows[8].Record.Scope <> 'StationA' OR "FRK_PersistImages".D001.Rows[8].Record.WriteKey <> 'degradationPercent' OR "FRK_PersistImages".D001.Rows[8].Record.Revision <> 1 OR "FRK_PersistImages".D001.Rows[8].Record.Kind <> 1 OR "FRK_PersistImages".D001.Rows[8].Record.ValueType <> 0 THEN RETURN; END_IF;
    #Ok := "FRK_ConfigDecode"(Text := STRING_TO_WSTRING("FRK_PersistImages".D001.Rows[8].Record.ValueText), Storage := 3, Minimum := 0.0, Maximum := 65535.0, MaxLength := 0, Value := "FRK_ConfigScratch".Value);
    IF NOT #Ok THEN RETURN; END_IF;
    IF NOT "FRK_PersistImages".D001.Rows[9].Used OR "FRK_PersistImages".D001.Rows[9].SchemaVersion <> 3 OR "FRK_PersistImages".D001.Rows[9].ModelCode <> '' OR "FRK_PersistImages".D001.Rows[9].Record.Scope <> 'StationA.Satellite' OR "FRK_PersistImages".D001.Rows[9].Record.WriteKey <> 'siteLabel' OR "FRK_PersistImages".D001.Rows[9].Record.Revision <> 1 OR "FRK_PersistImages".D001.Rows[9].Record.Kind <> 1 OR "FRK_PersistImages".D001.Rows[9].Record.ValueType <> 1 THEN RETURN; END_IF;
    #Ok := "FRK_ConfigDecode"(Text := STRING_TO_WSTRING("FRK_PersistImages".D001.Rows[9].Record.ValueText), Storage := 8, Minimum := 0.0, Maximum := 1.0, MaxLength := 80, Value := "FRK_ConfigScratch".Value);
    IF NOT #Ok THEN RETURN; END_IF;
    IF NOT "FRK_PersistImages".D001.Rows[10].Used OR "FRK_PersistImages".D001.Rows[10].SchemaVersion <> 3 OR "FRK_PersistImages".D001.Rows[10].ModelCode <> '' OR "FRK_PersistImages".D001.Rows[10].Record.Scope <> 'StationA.Satellite' OR "FRK_PersistImages".D001.Rows[10].Record.WriteKey <> 'enabled' OR "FRK_PersistImages".D001.Rows[10].Record.Revision <> 1 OR "FRK_PersistImages".D001.Rows[10].Record.Kind <> 1 OR "FRK_PersistImages".D001.Rows[10].Record.ValueType <> 2 THEN RETURN; END_IF;
    #Ok := "FRK_ConfigDecode"(Text := STRING_TO_WSTRING("FRK_PersistImages".D001.Rows[10].Record.ValueText), Storage := 1, Minimum := 0.0, Maximum := 1.0, MaxLength := 0, Value := "FRK_ConfigScratch".Value);
    IF NOT #Ok THEN RETURN; END_IF;
    IF NOT "FRK_PersistImages".D001.Rows[11].Used OR "FRK_PersistImages".D001.Rows[11].SchemaVersion <> 3 OR "FRK_PersistImages".D001.Rows[11].ModelCode <> '' OR "FRK_PersistImages".D001.Rows[11].Record.Scope <> 'StationA.Satellite' OR "FRK_PersistImages".D001.Rows[11].Record.WriteKey <> 'ratio' OR "FRK_PersistImages".D001.Rows[11].Record.Revision <> 1 OR "FRK_PersistImages".D001.Rows[11].Record.Kind <> 1 OR "FRK_PersistImages".D001.Rows[11].Record.ValueType <> 0 THEN RETURN; END_IF;
    #Ok := "FRK_ConfigDecode"(Text := STRING_TO_WSTRING("FRK_PersistImages".D001.Rows[11].Record.ValueText), Storage := 6, Minimum := -1000000.0, Maximum := 1000000.0, MaxLength := 0, Value := "FRK_ConfigScratch".Value);
    IF NOT #Ok THEN RETURN; END_IF;
    IF NOT "FRK_PersistImages".D001.Rows[12].Used OR "FRK_PersistImages".D001.Rows[12].SchemaVersion <> 3 OR "FRK_PersistImages".D001.Rows[12].ModelCode <> '' OR "FRK_PersistImages".D001.Rows[12].Record.Scope <> 'StationA.Satellite' OR "FRK_PersistImages".D001.Rows[12].Record.WriteKey <> 'gain' OR "FRK_PersistImages".D001.Rows[12].Record.Revision <> 1 OR "FRK_PersistImages".D001.Rows[12].Record.Kind <> 1 OR "FRK_PersistImages".D001.Rows[12].Record.ValueType <> 0 THEN RETURN; END_IF;
    #Ok := "FRK_ConfigDecode"(Text := STRING_TO_WSTRING("FRK_PersistImages".D001.Rows[12].Record.ValueText), Storage := 5, Minimum := -1000.0, Maximum := 1000.0, MaxLength := 0, Value := "FRK_ConfigScratch".Value);
    IF NOT #Ok THEN RETURN; END_IF;
    IF NOT "FRK_PersistImages".D001.Rows[13].Used OR "FRK_PersistImages".D001.Rows[13].SchemaVersion <> 3 OR "FRK_PersistImages".D001.Rows[13].ModelCode <> '' OR "FRK_PersistImages".D001.Rows[13].Record.Scope <> 'StationA.Satellite' OR "FRK_PersistImages".D001.Rows[13].Record.WriteKey <> 'grade' OR "FRK_PersistImages".D001.Rows[13].Record.Revision <> 1 OR "FRK_PersistImages".D001.Rows[13].Record.Kind <> 1 OR "FRK_PersistImages".D001.Rows[13].Record.ValueType <> 0 THEN RETURN; END_IF;
    #Ok := "FRK_ConfigDecode"(Text := STRING_TO_WSTRING("FRK_PersistImages".D001.Rows[13].Record.ValueText), Storage := 3, Minimum := 0.0, Maximum := 6.0, MaxLength := 0, Value := "FRK_ConfigScratch".Value);
    IF NOT #Ok THEN RETURN; END_IF;
    IF NOT "FRK_PersistImages".D001.Rows[14].Used OR "FRK_PersistImages".D001.Rows[14].SchemaVersion <> 3 OR "FRK_PersistImages".D001.Rows[14].ModelCode <> '' OR "FRK_PersistImages".D001.Rows[14].Record.Scope <> 'StationA.Satellite' OR "FRK_PersistImages".D001.Rows[14].Record.WriteKey <> 'offset.-1' OR "FRK_PersistImages".D001.Rows[14].Record.Revision <> 1 OR "FRK_PersistImages".D001.Rows[14].Record.Kind <> 1 OR "FRK_PersistImages".D001.Rows[14].Record.ValueType <> 0 THEN RETURN; END_IF;
    #Ok := "FRK_ConfigDecode"(Text := STRING_TO_WSTRING("FRK_PersistImages".D001.Rows[14].Record.ValueText), Storage := 2, Minimum := -32768.0, Maximum := 32767.0, MaxLength := 0, Value := "FRK_ConfigScratch".Value);
    IF NOT #Ok THEN RETURN; END_IF;
    IF NOT "FRK_PersistImages".D001.Rows[15].Used OR "FRK_PersistImages".D001.Rows[15].SchemaVersion <> 3 OR "FRK_PersistImages".D001.Rows[15].ModelCode <> '' OR "FRK_PersistImages".D001.Rows[15].Record.Scope <> 'StationA.Satellite' OR "FRK_PersistImages".D001.Rows[15].Record.WriteKey <> 'offset.0' OR "FRK_PersistImages".D001.Rows[15].Record.Revision <> 1 OR "FRK_PersistImages".D001.Rows[15].Record.Kind <> 1 OR "FRK_PersistImages".D001.Rows[15].Record.ValueType <> 0 THEN RETURN; END_IF;
    #Ok := "FRK_ConfigDecode"(Text := STRING_TO_WSTRING("FRK_PersistImages".D001.Rows[15].Record.ValueText), Storage := 2, Minimum := -32768.0, Maximum := 32767.0, MaxLength := 0, Value := "FRK_ConfigScratch".Value);
    IF NOT #Ok THEN RETURN; END_IF;
    IF NOT "FRK_PersistImages".D001.Rows[16].Used OR "FRK_PersistImages".D001.Rows[16].SchemaVersion <> 3 OR "FRK_PersistImages".D001.Rows[16].ModelCode <> '' OR "FRK_PersistImages".D001.Rows[16].Record.Scope <> 'StationA.Satellite' OR "FRK_PersistImages".D001.Rows[16].Record.WriteKey <> 'offset.1' OR "FRK_PersistImages".D001.Rows[16].Record.Revision <> 1 OR "FRK_PersistImages".D001.Rows[16].Record.Kind <> 1 OR "FRK_PersistImages".D001.Rows[16].Record.ValueType <> 0 THEN RETURN; END_IF;
    #Ok := "FRK_ConfigDecode"(Text := STRING_TO_WSTRING("FRK_PersistImages".D001.Rows[16].Record.ValueText), Storage := 2, Minimum := -32768.0, Maximum := 32767.0, MaxLength := 0, Value := "FRK_ConfigScratch".Value);
    IF NOT #Ok THEN RETURN; END_IF;
    IF NOT "FRK_PersistImages".D001.Rows[17].Used OR "FRK_PersistImages".D001.Rows[17].SchemaVersion <> 3 OR "FRK_PersistImages".D001.Rows[17].ModelCode <> '' OR "FRK_PersistImages".D001.Rows[17].Record.Scope <> 'StationA.Satellite' OR "FRK_PersistImages".D001.Rows[17].Record.WriteKey <> 'long.kkkkkkkkkkkkkkkkkkkkkkkkkkkkkkkkkkkkkkkkkkkkkkkkkkkkkkkkkkkkkkkkkkkkkkkkkkkkkkkkkkkkkkkkkkkkkkkkkkkkkkkkkkkkkkkkkkkkkkkkkkkkkkkkkkkkkkk' OR "FRK_PersistImages".D001.Rows[17].Record.Revision <> 1 OR "FRK_PersistImages".D001.Rows[17].Record.Kind <> 1 OR "FRK_PersistImages".D001.Rows[17].Record.ValueType <> 1 THEN RETURN; END_IF;
    #Ok := "FRK_ConfigDecode"(Text := STRING_TO_WSTRING("FRK_PersistImages".D001.Rows[17].Record.ValueText), Storage := 8, Minimum := 0.0, Maximum := 1.0, MaxLength := 80, Value := "FRK_ConfigScratch".Value);
    IF NOT #Ok THEN RETURN; END_IF;
    IF NOT "FRK_PersistImages".D001.Rows[18].Used OR "FRK_PersistImages".D001.Rows[18].SchemaVersion <> 3 OR "FRK_PersistImages".D001.Rows[18].ModelCode <> '' OR "FRK_PersistImages".D001.Rows[18].Record.Scope <> 'StationA.Satellite' OR "FRK_PersistImages".D001.Rows[18].Record.WriteKey <> 'small' OR "FRK_PersistImages".D001.Rows[18].Record.Revision <> 1 OR "FRK_PersistImages".D001.Rows[18].Record.Kind <> 1 OR "FRK_PersistImages".D001.Rows[18].Record.ValueType <> 0 THEN RETURN; END_IF;
    #Ok := "FRK_ConfigDecode"(Text := STRING_TO_WSTRING("FRK_PersistImages".D001.Rows[18].Record.ValueText), Storage := 3, Minimum := 0.0, Maximum := 255.0, MaxLength := 0, Value := "FRK_ConfigScratch".Value);
    IF NOT #Ok THEN RETURN; END_IF;
    IF NOT "FRK_PersistImages".D001.Rows[19].Used OR "FRK_PersistImages".D001.Rows[19].SchemaVersion <> 3 OR "FRK_PersistImages".D001.Rows[19].ModelCode <> '' OR "FRK_PersistImages".D001.Rows[19].Record.Scope <> 'StationA.Satellite.Inner' OR "FRK_PersistImages".D001.Rows[19].Record.WriteKey <> 'siteLabel' OR "FRK_PersistImages".D001.Rows[19].Record.Revision <> 1 OR "FRK_PersistImages".D001.Rows[19].Record.Kind <> 1 OR "FRK_PersistImages".D001.Rows[19].Record.ValueType <> 1 THEN RETURN; END_IF;
    #Ok := "FRK_ConfigDecode"(Text := STRING_TO_WSTRING("FRK_PersistImages".D001.Rows[19].Record.ValueText), Storage := 8, Minimum := 0.0, Maximum := 1.0, MaxLength := 80, Value := "FRK_ConfigScratch".Value);
    IF NOT #Ok THEN RETURN; END_IF;
    IF NOT "FRK_PersistImages".D001.Rows[20].Used OR "FRK_PersistImages".D001.Rows[20].SchemaVersion <> 3 OR "FRK_PersistImages".D001.Rows[20].ModelCode <> '' OR "FRK_PersistImages".D001.Rows[20].Record.Scope <> 'StationA.Satellite.Inner' OR "FRK_PersistImages".D001.Rows[20].Record.WriteKey <> 'enabled' OR "FRK_PersistImages".D001.Rows[20].Record.Revision <> 1 OR "FRK_PersistImages".D001.Rows[20].Record.Kind <> 1 OR "FRK_PersistImages".D001.Rows[20].Record.ValueType <> 2 THEN RETURN; END_IF;
    #Ok := "FRK_ConfigDecode"(Text := STRING_TO_WSTRING("FRK_PersistImages".D001.Rows[20].Record.ValueText), Storage := 1, Minimum := 0.0, Maximum := 1.0, MaxLength := 0, Value := "FRK_ConfigScratch".Value);
    IF NOT #Ok THEN RETURN; END_IF;
    IF NOT "FRK_PersistImages".D001.Rows[21].Used OR "FRK_PersistImages".D001.Rows[21].SchemaVersion <> 3 OR "FRK_PersistImages".D001.Rows[21].ModelCode <> '' OR "FRK_PersistImages".D001.Rows[21].Record.Scope <> 'StationA.Satellite.Inner' OR "FRK_PersistImages".D001.Rows[21].Record.WriteKey <> 'ratio' OR "FRK_PersistImages".D001.Rows[21].Record.Revision <> 1 OR "FRK_PersistImages".D001.Rows[21].Record.Kind <> 1 OR "FRK_PersistImages".D001.Rows[21].Record.ValueType <> 0 THEN RETURN; END_IF;
    #Ok := "FRK_ConfigDecode"(Text := STRING_TO_WSTRING("FRK_PersistImages".D001.Rows[21].Record.ValueText), Storage := 6, Minimum := -1000000.0, Maximum := 1000000.0, MaxLength := 0, Value := "FRK_ConfigScratch".Value);
    IF NOT #Ok THEN RETURN; END_IF;
    IF NOT "FRK_PersistImages".D001.Rows[22].Used OR "FRK_PersistImages".D001.Rows[22].SchemaVersion <> 3 OR "FRK_PersistImages".D001.Rows[22].ModelCode <> '' OR "FRK_PersistImages".D001.Rows[22].Record.Scope <> 'StationA.Satellite.Inner' OR "FRK_PersistImages".D001.Rows[22].Record.WriteKey <> 'gain' OR "FRK_PersistImages".D001.Rows[22].Record.Revision <> 1 OR "FRK_PersistImages".D001.Rows[22].Record.Kind <> 1 OR "FRK_PersistImages".D001.Rows[22].Record.ValueType <> 0 THEN RETURN; END_IF;
    #Ok := "FRK_ConfigDecode"(Text := STRING_TO_WSTRING("FRK_PersistImages".D001.Rows[22].Record.ValueText), Storage := 5, Minimum := -1000.0, Maximum := 1000.0, MaxLength := 0, Value := "FRK_ConfigScratch".Value);
    IF NOT #Ok THEN RETURN; END_IF;
    IF NOT "FRK_PersistImages".D001.Rows[23].Used OR "FRK_PersistImages".D001.Rows[23].SchemaVersion <> 3 OR "FRK_PersistImages".D001.Rows[23].ModelCode <> '' OR "FRK_PersistImages".D001.Rows[23].Record.Scope <> 'StationA.Satellite.Inner' OR "FRK_PersistImages".D001.Rows[23].Record.WriteKey <> 'grade' OR "FRK_PersistImages".D001.Rows[23].Record.Revision <> 1 OR "FRK_PersistImages".D001.Rows[23].Record.Kind <> 1 OR "FRK_PersistImages".D001.Rows[23].Record.ValueType <> 0 THEN RETURN; END_IF;
    #Ok := "FRK_ConfigDecode"(Text := STRING_TO_WSTRING("FRK_PersistImages".D001.Rows[23].Record.ValueText), Storage := 3, Minimum := 0.0, Maximum := 6.0, MaxLength := 0, Value := "FRK_ConfigScratch".Value);
    IF NOT #Ok THEN RETURN; END_IF;
    IF NOT "FRK_PersistImages".D001.Rows[24].Used OR "FRK_PersistImages".D001.Rows[24].SchemaVersion <> 3 OR "FRK_PersistImages".D001.Rows[24].ModelCode <> '' OR "FRK_PersistImages".D001.Rows[24].Record.Scope <> 'StationA.Satellite.Inner' OR "FRK_PersistImages".D001.Rows[24].Record.WriteKey <> 'offset.-1' OR "FRK_PersistImages".D001.Rows[24].Record.Revision <> 1 OR "FRK_PersistImages".D001.Rows[24].Record.Kind <> 1 OR "FRK_PersistImages".D001.Rows[24].Record.ValueType <> 0 THEN RETURN; END_IF;
    #Ok := "FRK_ConfigDecode"(Text := STRING_TO_WSTRING("FRK_PersistImages".D001.Rows[24].Record.ValueText), Storage := 2, Minimum := -32768.0, Maximum := 32767.0, MaxLength := 0, Value := "FRK_ConfigScratch".Value);
    IF NOT #Ok THEN RETURN; END_IF;
    IF NOT "FRK_PersistImages".D001.Rows[25].Used OR "FRK_PersistImages".D001.Rows[25].SchemaVersion <> 3 OR "FRK_PersistImages".D001.Rows[25].ModelCode <> '' OR "FRK_PersistImages".D001.Rows[25].Record.Scope <> 'StationA.Satellite.Inner' OR "FRK_PersistImages".D001.Rows[25].Record.WriteKey <> 'offset.0' OR "FRK_PersistImages".D001.Rows[25].Record.Revision <> 1 OR "FRK_PersistImages".D001.Rows[25].Record.Kind <> 1 OR "FRK_PersistImages".D001.Rows[25].Record.ValueType <> 0 THEN RETURN; END_IF;
    #Ok := "FRK_ConfigDecode"(Text := STRING_TO_WSTRING("FRK_PersistImages".D001.Rows[25].Record.ValueText), Storage := 2, Minimum := -32768.0, Maximum := 32767.0, MaxLength := 0, Value := "FRK_ConfigScratch".Value);
    IF NOT #Ok THEN RETURN; END_IF;
    IF NOT "FRK_PersistImages".D001.Rows[26].Used OR "FRK_PersistImages".D001.Rows[26].SchemaVersion <> 3 OR "FRK_PersistImages".D001.Rows[26].ModelCode <> '' OR "FRK_PersistImages".D001.Rows[26].Record.Scope <> 'StationA.Satellite.Inner' OR "FRK_PersistImages".D001.Rows[26].Record.WriteKey <> 'offset.1' OR "FRK_PersistImages".D001.Rows[26].Record.Revision <> 1 OR "FRK_PersistImages".D001.Rows[26].Record.Kind <> 1 OR "FRK_PersistImages".D001.Rows[26].Record.ValueType <> 0 THEN RETURN; END_IF;
    #Ok := "FRK_ConfigDecode"(Text := STRING_TO_WSTRING("FRK_PersistImages".D001.Rows[26].Record.ValueText), Storage := 2, Minimum := -32768.0, Maximum := 32767.0, MaxLength := 0, Value := "FRK_ConfigScratch".Value);
    IF NOT #Ok THEN RETURN; END_IF;
    IF NOT "FRK_PersistImages".D001.Rows[27].Used OR "FRK_PersistImages".D001.Rows[27].SchemaVersion <> 3 OR "FRK_PersistImages".D001.Rows[27].ModelCode <> '' OR "FRK_PersistImages".D001.Rows[27].Record.Scope <> 'StationA.Satellite.Inner' OR "FRK_PersistImages".D001.Rows[27].Record.WriteKey <> 'long.kkkkkkkkkkkkkkkkkkkkkkkkkkkkkkkkkkkkkkkkkkkkkkkkkkkkkkkkkkkkkkkkkkkkkkkkkkkkkkkkkkkkkkkkkkkkkkkkkkkkkkkkkkkkkkkkkkkkkkkkkkkkkkkkkkkkkkk' OR "FRK_PersistImages".D001.Rows[27].Record.Revision <> 1 OR "FRK_PersistImages".D001.Rows[27].Record.Kind <> 1 OR "FRK_PersistImages".D001.Rows[27].Record.ValueType <> 1 THEN RETURN; END_IF;
    #Ok := "FRK_ConfigDecode"(Text := STRING_TO_WSTRING("FRK_PersistImages".D001.Rows[27].Record.ValueText), Storage := 8, Minimum := 0.0, Maximum := 1.0, MaxLength := 80, Value := "FRK_ConfigScratch".Value);
    IF NOT #Ok THEN RETURN; END_IF;
    IF NOT "FRK_PersistImages".D001.Rows[28].Used OR "FRK_PersistImages".D001.Rows[28].SchemaVersion <> 3 OR "FRK_PersistImages".D001.Rows[28].ModelCode <> '' OR "FRK_PersistImages".D001.Rows[28].Record.Scope <> 'StationA.Satellite.Inner' OR "FRK_PersistImages".D001.Rows[28].Record.WriteKey <> 'small' OR "FRK_PersistImages".D001.Rows[28].Record.Revision <> 1 OR "FRK_PersistImages".D001.Rows[28].Record.Kind <> 1 OR "FRK_PersistImages".D001.Rows[28].Record.ValueType <> 0 THEN RETURN; END_IF;
    #Ok := "FRK_ConfigDecode"(Text := STRING_TO_WSTRING("FRK_PersistImages".D001.Rows[28].Record.ValueText), Storage := 3, Minimum := 0.0, Maximum := 255.0, MaxLength := 0, Value := "FRK_ConfigScratch".Value);
    IF NOT #Ok THEN RETURN; END_IF;
    #Stored := "FRK_ConfigFind"(Scope := 'StationA', Key := 'siteLabel', ModelCode := '');
    IF #Stored = 0 THEN
        FOR #Index := 1 TO 160 DO
            #Reserved := NOT "FRK_ConfigStore".Rows[#Index].Used;
            IF #Reserved THEN #Stored := #Index; EXIT; END_IF;
        END_FOR;
    END_IF;
    IF #Stored < 1 OR #Stored > 160 THEN RETURN; END_IF;
    #Targets[1] := #Stored;
    #Stored := "FRK_ConfigFind"(Scope := 'StationA', Key := 'enabled', ModelCode := '');
    IF #Stored = 0 THEN
        FOR #Index := 1 TO 160 DO
            #Reserved := NOT "FRK_ConfigStore".Rows[#Index].Used;
            FOR #Prior := 1 TO 1 DO IF #Targets[#Prior] = #Index THEN #Reserved := FALSE; END_IF; END_FOR;
            IF #Reserved THEN #Stored := #Index; EXIT; END_IF;
        END_FOR;
    END_IF;
    IF #Stored < 1 OR #Stored > 160 THEN RETURN; END_IF;
    #Targets[2] := #Stored;
    #Stored := "FRK_ConfigFind"(Scope := 'StationA', Key := 'ratio', ModelCode := '');
    IF #Stored = 0 THEN
        FOR #Index := 1 TO 160 DO
            #Reserved := NOT "FRK_ConfigStore".Rows[#Index].Used;
            FOR #Prior := 1 TO 2 DO IF #Targets[#Prior] = #Index THEN #Reserved := FALSE; END_IF; END_FOR;
            IF #Reserved THEN #Stored := #Index; EXIT; END_IF;
        END_FOR;
    END_IF;
    IF #Stored < 1 OR #Stored > 160 THEN RETURN; END_IF;
    #Targets[3] := #Stored;
    #Stored := "FRK_ConfigFind"(Scope := 'StationA', Key := 'gain', ModelCode := '');
    IF #Stored = 0 THEN
        FOR #Index := 1 TO 160 DO
            #Reserved := NOT "FRK_ConfigStore".Rows[#Index].Used;
            FOR #Prior := 1 TO 3 DO IF #Targets[#Prior] = #Index THEN #Reserved := FALSE; END_IF; END_FOR;
            IF #Reserved THEN #Stored := #Index; EXIT; END_IF;
        END_FOR;
    END_IF;
    IF #Stored < 1 OR #Stored > 160 THEN RETURN; END_IF;
    #Targets[4] := #Stored;
    #Stored := "FRK_ConfigFind"(Scope := 'StationA', Key := 'grade', ModelCode := '');
    IF #Stored = 0 THEN
        FOR #Index := 1 TO 160 DO
            #Reserved := NOT "FRK_ConfigStore".Rows[#Index].Used;
            FOR #Prior := 1 TO 4 DO IF #Targets[#Prior] = #Index THEN #Reserved := FALSE; END_IF; END_FOR;
            IF #Reserved THEN #Stored := #Index; EXIT; END_IF;
        END_FOR;
    END_IF;
    IF #Stored < 1 OR #Stored > 160 THEN RETURN; END_IF;
    #Targets[5] := #Stored;
    #Stored := "FRK_ConfigFind"(Scope := 'StationA', Key := 'small', ModelCode := '');
    IF #Stored = 0 THEN
        FOR #Index := 1 TO 160 DO
            #Reserved := NOT "FRK_ConfigStore".Rows[#Index].Used;
            FOR #Prior := 1 TO 5 DO IF #Targets[#Prior] = #Index THEN #Reserved := FALSE; END_IF; END_FOR;
            IF #Reserved THEN #Stored := #Index; EXIT; END_IF;
        END_FOR;
    END_IF;
    IF #Stored < 1 OR #Stored > 160 THEN RETURN; END_IF;
    #Targets[6] := #Stored;
    #Stored := "FRK_ConfigFind"(Scope := 'StationA', Key := 'long.kkkkkkkkkkkkkkkkkkkkkkkkkkkkkkkkkkkkkkkkkkkkkkkkkkkkkkkkkkkkkkkkkkkkkkkkkkkkkkkkkkkkkkkkkkkkkkkkkkkkkkkkkkkkkkkkkkkkkkkkkkkkkkkkkkkkkkk', ModelCode := '');
    IF #Stored = 0 THEN
        FOR #Index := 1 TO 160 DO
            #Reserved := NOT "FRK_ConfigStore".Rows[#Index].Used;
            FOR #Prior := 1 TO 6 DO IF #Targets[#Prior] = #Index THEN #Reserved := FALSE; END_IF; END_FOR;
            IF #Reserved THEN #Stored := #Index; EXIT; END_IF;
        END_FOR;
    END_IF;
    IF #Stored < 1 OR #Stored > 160 THEN RETURN; END_IF;
    #Targets[7] := #Stored;
    #Stored := "FRK_ConfigFind"(Scope := 'StationA', Key := 'degradationPercent', ModelCode := '');
    IF #Stored = 0 THEN
        FOR #Index := 1 TO 160 DO
            #Reserved := NOT "FRK_ConfigStore".Rows[#Index].Used;
